(* IEC 61131-3 sources: 2026_Projet_YGO_ExcavatriceDragage/TOOLS/TEST_AUTO_CI/RESULTS/M_MAIN/reports, 9 files *)

(* ---- FB_CfgT330Normalizer_test.st ---- *)
(* =======================================================================
   🧪 FB_CfgT330Normalizer — cas ST unitaires du plan T330 (C3 v1.3)
   ───────────────────────────────────────────────────────────────
   Périmètre STRICT : le FB de normalisation des réglages HAUT, en boîte
   noire (contrat light : Enable / InHoming -> Ready / Corrected).
   Aucune assertion ne porte sur un consommateur (PRG_03 / PRG_04 /
   PRG_06 / GVL_PERSISTENT) : ces cas relèvent d'un lot d'intégration
   dédié (voir TASK_CONTRACT_T341, section « hors scope »).

   ── Conventions ───────────────────────────────────────────────────────
   1) 1 appel fb(...) = 1 scan.
   2) ⚠️ STruCpp v0.6.2 passe les VAR_IN_OUT par COPIE et ne génère que le
      copy-IN. La restitution `cfg := fb.CommunCfg;` est donc OBLIGATOIRE
      après chaque appel : elle émule la sémantique par RÉFÉRENCE de
      CODESYS. Sans elle, toute assertion de correction serait VACUE
      (le FB écrirait dans sa copie privée, jamais dans la variable de test).
      Le post-traitement `inject_var_in_out_copyout.py` ne s'applique PAS à
      une VAR déclarée dans un bloc `VAR` local de TEST (sa regex exige le
      préfixe `s.` que ce build n'émet pas) — d'où l'émulation explicite.
   3) ⚠️ Aucune assertion n'est placée dans une boucle FOR/WHILE : ce build
      STruCpp SUPPRIME silencieusement les ASSERT_* du corps d'une boucle
      (vérifié dans le C++ généré). Les balayages sont donc déroulés.
   4) Tolérance 1e-6 : les REAL sont en simple précision, un littéral ST est
      lu en double — un écart de ~1,4e-7 est normal sur 7,4999.
   5) Amorcage : le FB amorce ses mémoires de front au PREMIER scan où
      `Enable` est vrai, depuis les valeurs RESTAURÉES (piège P2 du cadrage).
      Une stimulation « saisie opérateur » se joue donc au scan SUIVANT.

   Référence : DOC/WFLOW/AUDITS/DESIGN/PLAN_T330_C3_INVARIANT_HAUT_v1.0.md §4.2
   ======================================================================= *)

SETUP
VAR
    FB       : FB_CfgT330Normalizer;
    WinchCfg : ST_WinchCfg;
    ComCfg   : ST_CommunCfg;
END_VAR
END_SETUP

(* ── Groupe A · Normalisation (TC-P10-056 .. TC-P10-062) ──────────────── *)

TEST 'TC-P10-056 R1 — FDC saisi trop haut : FDC corrige, TOP preserve'
VAR
    winchCfg  : ST_WinchCfg;
    communCfg : ST_CommunCfg;
END_VAR
    (* Scan 1 : amorcage sur la config restauree valide (8,50 / 7,50 / 0,50). *)
    winchCfg.CfgTopSensorPos_M := 8.5;
    communCfg.CfgCableLimitAscent_M := 7.5;
    communCfg.WinchSlowdownDistanceTop_M := 0.5;
    FB.Enable := TRUE;
    FB.InHoming := FALSE;
    FB(WinchCfgM1 := winchCfg, CommunCfg := communCfg);
    winchCfg := FB.WinchCfgM1;  communCfg := FB.CommunCfg;
    ASSERT_FALSE(FB.Corrected, 'Scan d amorcage : config valide, aucune correction');

    (* Scan 2 : l'operateur saisit FDC = 8,70 m (TOP inchange a 8,50 m). *)
    communCfg.CfgCableLimitAscent_M := 8.7;
    FB(WinchCfgM1 := winchCfg, CommunCfg := communCfg);
    winchCfg := FB.WinchCfgM1;  communCfg := FB.CommunCfg;
    ASSERT_NEAR(communCfg.CfgCableLimitAscent_M, 7.5, 0.000001,
                'R1 : FDC ramene a TOP - 1,00 m = 7,50');
    ASSERT_NEAR(winchCfg.CfgTopSensorPos_M, 8.5, 0.000001, 'R1 : le TOP n est PAS modifie');
    ASSERT_TRUE(FB.Corrected, 'R1 : une correction a eu lieu, message emis');
END_TEST

TEST 'TC-P10-057 R2 — TOP saisi trop bas : TOP corrige, FDC preserve'
VAR
    winchCfg  : ST_WinchCfg;
    communCfg : ST_CommunCfg;
END_VAR
    winchCfg.CfgTopSensorPos_M := 8.5;
    communCfg.CfgCableLimitAscent_M := 7.5;
    communCfg.WinchSlowdownDistanceTop_M := 0.5;
    FB.Enable := TRUE;
    FB.InHoming := FALSE;
    FB(WinchCfgM1 := winchCfg, CommunCfg := communCfg);
    winchCfg := FB.WinchCfgM1;  communCfg := FB.CommunCfg;

    (* Scan 2 : l'operateur saisit TOP = 7,00 m (FDC inchange a 7,50 m). *)
    winchCfg.CfgTopSensorPos_M := 7.0;
    FB(WinchCfgM1 := winchCfg, CommunCfg := communCfg);
    winchCfg := FB.WinchCfgM1;  communCfg := FB.CommunCfg;
    ASSERT_NEAR(winchCfg.CfgTopSensorPos_M, 8.5, 0.000001,
                'R2 : TOP ramene a FDC + 1,00 m = 8,50 (le champ saisi est corrige)');
    ASSERT_NEAR(communCfg.CfgCableLimitAscent_M, 7.5, 0.000001, 'R2 : le FDC n est PAS modifie');
    ASSERT_TRUE(FB.Corrected, 'R2 : une correction a eu lieu, message emis');
END_TEST

TEST 'TC-P10-058 R1 — Delta = 0,90 m : correction du champ saisi (FDC)'
VAR
    winchCfg  : ST_WinchCfg;
    communCfg : ST_CommunCfg;
END_VAR
    winchCfg.CfgTopSensorPos_M := 8.5;
    communCfg.CfgCableLimitAscent_M := 7.5;
    communCfg.WinchSlowdownDistanceTop_M := 0.5;
    FB.Enable := TRUE;
    FB.InHoming := FALSE;
    FB(WinchCfgM1 := winchCfg, CommunCfg := communCfg);
    winchCfg := FB.WinchCfgM1;  communCfg := FB.CommunCfg;

    (* Scan 2 : FDC = 7,60 m => Delta = 8,50 - 7,60 = 0,90 m < 1,00 m. *)
    communCfg.CfgCableLimitAscent_M := 7.6;
    FB(WinchCfgM1 := winchCfg, CommunCfg := communCfg);
    winchCfg := FB.WinchCfgM1;  communCfg := FB.CommunCfg;
    ASSERT_NEAR(communCfg.CfgCableLimitAscent_M, 7.5, 0.000001, 'Delta < 1,00 m : FDC ramene a 7,50');
    ASSERT_NEAR(winchCfg.CfgTopSensorPos_M, 8.5, 0.000001, 'Delta < 1,00 m : TOP preserve');
    ASSERT_TRUE(FB.Corrected, 'Delta < 1,00 m : correction signalee');
END_TEST

TEST 'TC-P10-059 R3 — plancher du ralentissement haut (0,20 -> 0,50)'
VAR
    winchCfg  : ST_WinchCfg;
    communCfg : ST_CommunCfg;
END_VAR
    winchCfg.CfgTopSensorPos_M := 8.5;
    communCfg.CfgCableLimitAscent_M := 7.5;
    communCfg.WinchSlowdownDistanceTop_M := 0.5;
    FB.Enable := TRUE;
    FB.InHoming := FALSE;
    FB(WinchCfgM1 := winchCfg, CommunCfg := communCfg);
    winchCfg := FB.WinchCfgM1;  communCfg := FB.CommunCfg;

    (* Scan 2 : ralentissement saisi a 0,20 m (< 0,50 m). *)
    communCfg.WinchSlowdownDistanceTop_M := 0.2;
    FB(WinchCfgM1 := winchCfg, CommunCfg := communCfg);
    winchCfg := FB.WinchCfgM1;  communCfg := FB.CommunCfg;
    ASSERT_NEAR(communCfg.WinchSlowdownDistanceTop_M, 0.5, 0.000001,
                'R3 : ralentissement ramene au plancher 0,50 m');
    ASSERT_NEAR(winchCfg.CfgTopSensorPos_M, 8.5, 0.000001, 'R3 : TOP inchange');
    ASSERT_NEAR(communCfg.CfgCableLimitAscent_M, 7.5, 0.000001, 'R3 : FDC inchange');
    ASSERT_TRUE(FB.Corrected, 'R3 : correction signalee');
END_TEST

TEST 'TC-P10-060 config valide (Delta = 2,50) : aucune correction, aucun message'
VAR
    winchCfg  : ST_WinchCfg;
    communCfg : ST_CommunCfg;
END_VAR
    winchCfg.CfgTopSensorPos_M := 8.5;
    communCfg.CfgCableLimitAscent_M := 7.5;
    communCfg.WinchSlowdownDistanceTop_M := 0.5;
    FB.Enable := TRUE;
    FB.InHoming := FALSE;
    FB(WinchCfgM1 := winchCfg, CommunCfg := communCfg);
    winchCfg := FB.WinchCfgM1;  communCfg := FB.CommunCfg;

    (* Scan 2 : TOP = 10,00 m, FDC = 7,50 m => Delta = 2,50 m, valide. *)
    winchCfg.CfgTopSensorPos_M := 10.0;
    FB(WinchCfgM1 := winchCfg, CommunCfg := communCfg);
    winchCfg := FB.WinchCfgM1;  communCfg := FB.CommunCfg;
    ASSERT_NEAR(winchCfg.CfgTopSensorPos_M, 10.0, 0.000001, 'Config valide : TOP preserve');
    ASSERT_NEAR(communCfg.CfgCableLimitAscent_M, 7.5, 0.000001, 'Config valide : FDC preserve');
    ASSERT_FALSE(FB.Corrected, 'Config valide : AUCUN message (compteur de messages = 0)');
END_TEST

TEST 'TC-P10-061 Q17 — les DEUX champs changent au meme scan : TOP preserve, FDC corrige'
VAR
    winchCfg  : ST_WinchCfg;
    communCfg : ST_CommunCfg;
END_VAR
    winchCfg.CfgTopSensorPos_M := 8.5;
    communCfg.CfgCableLimitAscent_M := 7.5;
    communCfg.WinchSlowdownDistanceTop_M := 0.5;
    FB.Enable := TRUE;
    FB.InHoming := FALSE;
    FB(WinchCfgM1 := winchCfg, CommunCfg := communCfg);
    winchCfg := FB.WinchCfgM1;  communCfg := FB.CommunCfg;

    (* Scan 2 : les 3 reglages changent ensemble : FDC 9,50 / TOP 8,00 / slowdown 0,10. *)
    communCfg.CfgCableLimitAscent_M := 9.5;
    winchCfg.CfgTopSensorPos_M := 8.0;
    communCfg.WinchSlowdownDistanceTop_M := 0.1;
    FB(WinchCfgM1 := winchCfg, CommunCfg := communCfg);
    winchCfg := FB.WinchCfgM1;  communCfg := FB.CommunCfg;
    ASSERT_NEAR(winchCfg.CfgTopSensorPos_M, 8.0, 0.000001, 'Q17 : le TOP saisi est PRESERVE');
    ASSERT_NEAR(communCfg.CfgCableLimitAscent_M, 7.0, 0.000001,
                'Q17 : FDC = TOP - 1,00 m = 7,00 (R0 a d abord ramene 9,50 a 9,00)');
    ASSERT_NEAR(communCfg.WinchSlowdownDistanceTop_M, 0.5, 0.000001, 'R3 : ralentissement ramene a 0,50');
    ASSERT_TRUE(FB.Corrected, 'Q17 : les trois corrections sont signalees');
END_TEST

TEST 'TC-P10-062 FDC = 0,00 m (borne basse, Delta valide) : accepte, aucune correction'
VAR
    winchCfg  : ST_WinchCfg;
    communCfg : ST_CommunCfg;
END_VAR
    winchCfg.CfgTopSensorPos_M := 8.5;
    communCfg.CfgCableLimitAscent_M := 7.5;
    communCfg.WinchSlowdownDistanceTop_M := 0.5;
    FB.Enable := TRUE;
    FB.InHoming := FALSE;
    FB(WinchCfgM1 := winchCfg, CommunCfg := communCfg);
    winchCfg := FB.WinchCfgM1;  communCfg := FB.CommunCfg;

    (* Scan 2 : FDC = 0,00 m => Delta = 8,50 m, valide. La borne basse est INCLUSE. *)
    communCfg.CfgCableLimitAscent_M := 0.0;
    FB(WinchCfgM1 := winchCfg, CommunCfg := communCfg);
    winchCfg := FB.WinchCfgM1;  communCfg := FB.CommunCfg;
    ASSERT_NEAR(communCfg.CfgCableLimitAscent_M, 0.0, 0.000001,
                'FDC a la borne basse : valeur ACCEPTEE telle quelle');
    ASSERT_NEAR(winchCfg.CfgTopSensorPos_M, 8.5, 0.000001, 'FDC a la borne basse : TOP inchange');
    ASSERT_FALSE(FB.Corrected, 'FDC a la borne basse : aucune correction, aucun message');
END_TEST

(* ── Groupe B · Idempotence et non-rebond (TC-P10-063 .. TC-P10-068) ──── *)

TEST 'TC-P10-063 Q24 — idempotence : le 2e scan apres correction ne corrige PLUS'
VAR
    winchCfg  : ST_WinchCfg;
    communCfg : ST_CommunCfg;
END_VAR
    winchCfg.CfgTopSensorPos_M := 8.5;
    communCfg.CfgCableLimitAscent_M := 7.5;
    communCfg.WinchSlowdownDistanceTop_M := 0.5;
    FB.Enable := TRUE;
    FB.InHoming := FALSE;
    FB(WinchCfgM1 := winchCfg, CommunCfg := communCfg);
    winchCfg := FB.WinchCfgM1;  communCfg := FB.CommunCfg;

    (* Scan 2 : correction (FDC 8,70 -> 7,50). *)
    communCfg.CfgCableLimitAscent_M := 8.7;
    FB(WinchCfgM1 := winchCfg, CommunCfg := communCfg);
    winchCfg := FB.WinchCfgM1;  communCfg := FB.CommunCfg;
    ASSERT_NEAR(communCfg.CfgCableLimitAscent_M, 7.5, 0.000001, 'Scan 2 : FDC corrige a 7,50');

    (* Scan 3 : rejeu SANS nouvelle saisie => ni correction, ni message, valeur stable. *)
    FB(WinchCfgM1 := winchCfg, CommunCfg := communCfg);
    winchCfg := FB.WinchCfgM1;  communCfg := FB.CommunCfg;
    ASSERT_NEAR(communCfg.CfgCableLimitAscent_M, 7.5, 0.000001, 'Scan 3 : valeur STABLE a 7,50');
    ASSERT_FALSE(FB.Corrected, 'Scan 3 : AUCUNE seconde correction (test probatoire de Q24)');
END_TEST

TEST 'TC-P10-064 reserve EXACTEMENT 1,00 m : aucune correction (aucun epsilon)'
VAR
    winchCfg  : ST_WinchCfg;
    communCfg : ST_CommunCfg;
END_VAR
    winchCfg.CfgTopSensorPos_M := 8.5;
    communCfg.CfgCableLimitAscent_M := 7.5;
    communCfg.WinchSlowdownDistanceTop_M := 0.5;
    FB.Enable := TRUE;
    FB.InHoming := FALSE;
    FB(WinchCfgM1 := winchCfg, CommunCfg := communCfg);
    winchCfg := FB.WinchCfgM1;  communCfg := FB.CommunCfg;
    ASSERT_FALSE(FB.Corrected, 'Delta = 1,00 m exactement : aucune correction (comparaison stricte)');
    ASSERT_NEAR(winchCfg.CfgTopSensorPos_M - communCfg.CfgCableLimitAscent_M, 1.0, 0.000001,
                'Le flottant est EXACT : 8,50 - 7,50 = 1,00 (aucun eps necessaire)');

    (* Scan 2 : rejeu identique — la reserve reste exactement 1,00 m. *)
    FB(WinchCfgM1 := winchCfg, CommunCfg := communCfg);
    winchCfg := FB.WinchCfgM1;  communCfg := FB.CommunCfg;
    ASSERT_FALSE(FB.Corrected, 'Scan 2 : aucune oscillation autour du seuil');
END_TEST

TEST 'TC-P10-065 pt1 balayage 7,4999 — Delta = 1,0001 m : FDC conserve'
VAR
    winchCfg  : ST_WinchCfg;
    communCfg : ST_CommunCfg;
END_VAR
    winchCfg.CfgTopSensorPos_M := 8.5;
    communCfg.CfgCableLimitAscent_M := 7.5;
    communCfg.WinchSlowdownDistanceTop_M := 0.5;
    FB.Enable := TRUE;
    FB.InHoming := FALSE;
    FB(WinchCfgM1 := winchCfg, CommunCfg := communCfg);
    winchCfg := FB.WinchCfgM1;  communCfg := FB.CommunCfg;

    communCfg.CfgCableLimitAscent_M := 7.4999;
    FB(WinchCfgM1 := winchCfg, CommunCfg := communCfg);
    winchCfg := FB.WinchCfgM1;  communCfg := FB.CommunCfg;
    ASSERT_NEAR(communCfg.CfgCableLimitAscent_M, 7.4999, 0.000001,
                'Delta > 1,00 m : FDC conserve tel quel');
    ASSERT_FALSE(FB.Corrected, 'Delta > 1,00 m : aucun message');
END_TEST

TEST 'TC-P10-065 pt2 balayage 7,5000 — Delta = 1,00 m exactement : FDC conserve'
VAR
    winchCfg  : ST_WinchCfg;
    communCfg : ST_CommunCfg;
END_VAR
    winchCfg.CfgTopSensorPos_M := 8.5;
    communCfg.CfgCableLimitAscent_M := 7.5;
    communCfg.WinchSlowdownDistanceTop_M := 0.5;
    FB.Enable := TRUE;
    FB.InHoming := FALSE;
    FB(WinchCfgM1 := winchCfg, CommunCfg := communCfg);
    winchCfg := FB.WinchCfgM1;  communCfg := FB.CommunCfg;

    communCfg.CfgCableLimitAscent_M := 7.5;
    FB(WinchCfgM1 := winchCfg, CommunCfg := communCfg);
    winchCfg := FB.WinchCfgM1;  communCfg := FB.CommunCfg;
    ASSERT_NEAR(communCfg.CfgCableLimitAscent_M, 7.5, 0.000001,
                'Delta = 1,00 m (point limite INCLUS) : FDC conserve');
    ASSERT_FALSE(FB.Corrected, 'Delta = 1,00 m : aucun message');
END_TEST

TEST 'TC-P10-065 pt3 balayage 7,5001 — Delta = 0,9999 m : FDC corrige, une seule fois'
VAR
    winchCfg  : ST_WinchCfg;
    communCfg : ST_CommunCfg;
END_VAR
    winchCfg.CfgTopSensorPos_M := 8.5;
    communCfg.CfgCableLimitAscent_M := 7.5;
    communCfg.WinchSlowdownDistanceTop_M := 0.5;
    FB.Enable := TRUE;
    FB.InHoming := FALSE;
    FB(WinchCfgM1 := winchCfg, CommunCfg := communCfg);
    winchCfg := FB.WinchCfgM1;  communCfg := FB.CommunCfg;

    communCfg.CfgCableLimitAscent_M := 7.5001;
    FB(WinchCfgM1 := winchCfg, CommunCfg := communCfg);
    winchCfg := FB.WinchCfgM1;  communCfg := FB.CommunCfg;
    ASSERT_NEAR(communCfg.CfgCableLimitAscent_M, 7.5, 0.000001, 'Delta < 1,00 m : FDC ramene a 7,50');
    ASSERT_TRUE(FB.Corrected, 'Delta < 1,00 m : correction signalee');

    (* Scan suivant : la valeur corrigee ne rebondit pas (aucune oscillation au seuil). *)
    FB(WinchCfgM1 := winchCfg, CommunCfg := communCfg);
    winchCfg := FB.WinchCfgM1;  communCfg := FB.CommunCfg;
    ASSERT_FALSE(FB.Corrected, 'Scan suivant : aucune seconde correction (pas d oscillation)');
END_TEST

TEST 'TC-P10-066 LIMITE DECLAREE — guerre d ecriture IHM : correction a CHAQUE scan'
VAR
    winchCfg  : ST_WinchCfg;
    communCfg : ST_CommunCfg;
END_VAR
    (* ⚠️ Ce cas fige une LIMITE ASSUMEE du lot (plan v1.3 §4.2, C3), PAS une exigence :
       si le panneau IHM reecrit 8,70 m a CHAQUE scan, la normalisation corrige a chaque
       scan et le message rebondit — aucun amortissement n'est specifie ni implemente.
       Le test est volontairement falsifiable : ajouter un anti-rebond le fera echouer,
       ce qui forcera une decision DOCUMENTEE plutot qu'une derive silencieuse.
       Balayage DEROULE (3 scans) : une assertion dans une boucle serait supprimee
       silencieusement par STruCpp et le test deviendrait VACUE. *)
    winchCfg.CfgTopSensorPos_M := 8.5;
    communCfg.CfgCableLimitAscent_M := 7.5;
    communCfg.WinchSlowdownDistanceTop_M := 0.5;
    FB.Enable := TRUE;
    FB.InHoming := FALSE;
    FB(WinchCfgM1 := winchCfg, CommunCfg := communCfg);
    winchCfg := FB.WinchCfgM1;  communCfg := FB.CommunCfg;

    (* Scan 2. *)
    communCfg.CfgCableLimitAscent_M := 8.7;
    FB(WinchCfgM1 := winchCfg, CommunCfg := communCfg);
    winchCfg := FB.WinchCfgM1;  communCfg := FB.CommunCfg;
    ASSERT_NEAR(communCfg.CfgCableLimitAscent_M, 7.5, 0.000001, 'Scan 2 : correction reappliquee');
    ASSERT_TRUE(FB.Corrected, 'Scan 2 : message emis (rebond ASSUME)');

    (* Scan 3. *)
    communCfg.CfgCableLimitAscent_M := 8.7;
    FB(WinchCfgM1 := winchCfg, CommunCfg := communCfg);
    winchCfg := FB.WinchCfgM1;  communCfg := FB.CommunCfg;
    ASSERT_NEAR(communCfg.CfgCableLimitAscent_M, 7.5, 0.000001, 'Scan 3 : correction reappliquee');
    ASSERT_TRUE(FB.Corrected, 'Scan 3 : message emis (rebond ASSUME)');

    (* Scan 4. *)
    communCfg.CfgCableLimitAscent_M := 8.7;
    FB(WinchCfgM1 := winchCfg, CommunCfg := communCfg);
    winchCfg := FB.WinchCfgM1;  communCfg := FB.CommunCfg;
    ASSERT_NEAR(communCfg.CfgCableLimitAscent_M, 7.5, 0.000001, 'Scan 4 : correction reappliquee');
    ASSERT_TRUE(FB.Corrected, 'Scan 4 : message emis (rebond ASSUME)');
END_TEST

TEST 'TC-P10-067 valeur IDENTIQUE re-saisie : aucun front, aucune correction'
VAR
    winchCfg  : ST_WinchCfg;
    communCfg : ST_CommunCfg;
END_VAR
    winchCfg.CfgTopSensorPos_M := 8.5;
    communCfg.CfgCableLimitAscent_M := 7.5;
    communCfg.WinchSlowdownDistanceTop_M := 0.5;
    FB.Enable := TRUE;
    FB.InHoming := FALSE;
    FB(WinchCfgM1 := winchCfg, CommunCfg := communCfg);
    winchCfg := FB.WinchCfgM1;  communCfg := FB.CommunCfg;

    (* Scan 2 : le champ est REEcrit avec la MEME valeur (8,50 -> 8,50). *)
    winchCfg.CfgTopSensorPos_M := 8.5;
    FB(WinchCfgM1 := winchCfg, CommunCfg := communCfg);
    winchCfg := FB.WinchCfgM1;  communCfg := FB.CommunCfg;
    ASSERT_FALSE(FB.Corrected, 'Valeur identique re-saisie : aucun front, aucun message');
    ASSERT_NEAR(winchCfg.CfgTopSensorPos_M, 8.5, 0.000001, 'Valeur identique : TOP inchange');
END_TEST

TEST 'TC-P10-068 changement de page IHM sans modification : aucune correction'
VAR
    winchCfg  : ST_WinchCfg;
    communCfg : ST_CommunCfg;
END_VAR
    winchCfg.CfgTopSensorPos_M := 8.5;
    communCfg.CfgCableLimitAscent_M := 7.5;
    communCfg.WinchSlowdownDistanceTop_M := 0.5;
    FB.Enable := TRUE;
    FB.InHoming := FALSE;
    FB(WinchCfgM1 := winchCfg, CommunCfg := communCfg);
    winchCfg := FB.WinchCfgM1;  communCfg := FB.CommunCfg;

    (* Scan 2 : page quittee => normalisation suspendue, AUCUNE valeur modifiee. *)
    FB.Enable := FALSE;
    FB(WinchCfgM1 := winchCfg, CommunCfg := communCfg);
    winchCfg := FB.WinchCfgM1;  communCfg := FB.CommunCfg;
    ASSERT_FALSE(FB.Corrected, 'Normalisation suspendue : aucun message');
    ASSERT_FALSE(FB.Ready, 'Normalisation suspendue : Ready = FALSE');

    (* Scan 3 : retour sur la page, valeurs inchangees => ni front, ni correction. *)
    FB.Enable := TRUE;
    FB(WinchCfgM1 := winchCfg, CommunCfg := communCfg);
    winchCfg := FB.WinchCfgM1;  communCfg := FB.CommunCfg;
    ASSERT_FALSE(FB.Corrected, 'Retour de page sans modification : aucune correction');
    ASSERT_NEAR(winchCfg.CfgTopSensorPos_M, 8.5, 0.000001, 'Retour de page : TOP inchange');
    ASSERT_NEAR(communCfg.CfgCableLimitAscent_M, 7.5, 0.000001, 'Retour de page : FDC inchange');
END_TEST

(* ── Groupe C · Boot, restauration, hot restart (TC-P10-069 .. TC-P10-074) ─ *)

TEST 'TC-P10-069 NVRAM valide au demarrage a froid : 0 correction, valeurs preservees'
VAR
    winchCfg  : ST_WinchCfg;
    communCfg : ST_CommunCfg;
END_VAR
    winchCfg.CfgTopSensorPos_M := 8.5;
    communCfg.CfgCableLimitAscent_M := 7.5;
    communCfg.WinchSlowdownDistanceTop_M := 0.5;
    FB.Enable := TRUE;
    FB.InHoming := FALSE;
    FB(WinchCfgM1 := winchCfg, CommunCfg := communCfg);
    winchCfg := FB.WinchCfgM1;  communCfg := FB.CommunCfg;
    ASSERT_TRUE(FB.Ready, 'Normalisation ARMED des le premier scan apres restauration');
    ASSERT_FALSE(FB.Corrected, 'NVRAM valide : aucune correction');
    ASSERT_NEAR(winchCfg.CfgTopSensorPos_M, 8.5, 0.000001, 'NVRAM valide : TOP preserve');
    ASSERT_NEAR(communCfg.CfgCableLimitAscent_M, 7.5, 0.000001, 'NVRAM valide : FDC preserve');
    ASSERT_NEAR(communCfg.WinchSlowdownDistanceTop_M, 0.5, 0.000001, 'NVRAM valide : ralentissement preserve');
END_TEST

TEST 'TC-P10-070 NVRAM invalide au demarrage a froid : Q17 (TOP preserve, FDC corrige)'
VAR
    winchCfg  : ST_WinchCfg;
    communCfg : ST_CommunCfg;
END_VAR
    (* NVRAM restauree INVALIDE : TOP = 7,00 m / FDC = 7,50 m. *)
    winchCfg.CfgTopSensorPos_M := 7.0;
    communCfg.CfgCableLimitAscent_M := 7.5;
    communCfg.WinchSlowdownDistanceTop_M := 0.5;
    FB.Enable := TRUE;
    FB.InHoming := FALSE;
    FB(WinchCfgM1 := winchCfg, CommunCfg := communCfg);
    winchCfg := FB.WinchCfgM1;  communCfg := FB.CommunCfg;
    ASSERT_NEAR(winchCfg.CfgTopSensorPos_M, 7.0, 0.000001,
                'Q17 : le TOP restaure est PRESERVE (c est la cote gravee par le homing)');
    ASSERT_NEAR(communCfg.CfgCableLimitAscent_M, 6.0, 0.000001, 'Q17 : FDC = TOP - 1,00 m = 6,00');
    ASSERT_TRUE(FB.Corrected, 'NVRAM invalide : correction signalee');
END_TEST

TEST 'TC-P10-071 premier scan NOT Initialized : normalisation INHIBEE, aucune ecriture'
VAR
    winchCfg  : ST_WinchCfg;
    communCfg : ST_CommunCfg;
END_VAR
    (* Ponts non restaures : les valeurs presentes sont les DEFAUTS DUT, pas une saisie. *)
    winchCfg.CfgTopSensorPos_M := 99.0;
    communCfg.CfgCableLimitAscent_M := 99.0;
    communCfg.WinchSlowdownDistanceTop_M := 99.0;
    FB.Enable := FALSE;
    FB.InHoming := FALSE;
    FB(WinchCfgM1 := winchCfg, CommunCfg := communCfg);
    winchCfg := FB.WinchCfgM1;  communCfg := FB.CommunCfg;
    ASSERT_FALSE(FB.Ready, 'NOT Initialized : normalisation NON armee');
    ASSERT_FALSE(FB.Corrected, 'NOT Initialized : aucun message');
    ASSERT_NEAR(winchCfg.CfgTopSensorPos_M, 99.0, 0.000001, 'NOT Initialized : AUCUNE ecriture TOP');
    ASSERT_NEAR(communCfg.CfgCableLimitAscent_M, 99.0, 0.000001, 'NOT Initialized : AUCUNE ecriture FDC');
    ASSERT_NEAR(communCfg.WinchSlowdownDistanceTop_M, 99.0, 0.000001,
                'NOT Initialized : AUCUNE ecriture ralentissement');
END_TEST

TEST 'TC-P10-074 ptA restauration NVRAM : AUCUNE correction fantome (defauts DUT -> restaure)'
VAR
    winchCfg  : ST_WinchCfg;
    communCfg : ST_CommunCfg;
END_VAR
    (* PREUVE EXIGEE par le plan §2.2 point 3 : la transition « defauts DUT ->
       valeurs RESTAUREES » ne doit PAS etre prise pour une saisie operateur. *)
    winchCfg.CfgTopSensorPos_M := 8.5;      (* defauts DUT au 1er scan *)
    communCfg.CfgCableLimitAscent_M := 7.5;
    communCfg.WinchSlowdownDistanceTop_M := 0.5;
    FB.Enable := FALSE;                     (* ponts non restaures *)
    FB.InHoming := FALSE;
    FB(WinchCfgM1 := winchCfg, CommunCfg := communCfg);
    winchCfg := FB.WinchCfgM1;  communCfg := FB.CommunCfg;

    winchCfg.CfgTopSensorPos_M := 8.5;      (* valeurs RESTAUREES, valides *)
    communCfg.CfgCableLimitAscent_M := 7.5;
    communCfg.WinchSlowdownDistanceTop_M := 0.5;
    FB.Enable := TRUE;
    FB(WinchCfgM1 := winchCfg, CommunCfg := communCfg);
    winchCfg := FB.WinchCfgM1;  communCfg := FB.CommunCfg;
    ASSERT_FALSE(FB.Corrected, 'Restauration NVRAM : AUCUNE correction fantome');
    ASSERT_NEAR(winchCfg.CfgTopSensorPos_M, 8.5, 0.000001, 'Restauration NVRAM : TOP preserve');
    ASSERT_NEAR(communCfg.CfgCableLimitAscent_M, 7.5, 0.000001, 'Restauration NVRAM : FDC preserve');
END_TEST

TEST 'TC-P10-074 ptB download/RTS : comportement DETERMINISTE, une seule correction'
VAR
    winchCfg  : ST_WinchCfg;
    communCfg : ST_CommunCfg;
END_VAR
    (* NVRAM restauree INVALIDE apres download : une correction, jamais repetee. *)
    winchCfg.CfgTopSensorPos_M := 7.0;
    communCfg.CfgCableLimitAscent_M := 7.5;
    communCfg.WinchSlowdownDistanceTop_M := 0.5;
    FB.Enable := TRUE;
    FB.InHoming := FALSE;
    FB(WinchCfgM1 := winchCfg, CommunCfg := communCfg);
    winchCfg := FB.WinchCfgM1;  communCfg := FB.CommunCfg;
    ASSERT_TRUE(FB.Corrected, 'NVRAM invalide : une correction, signalee');
    ASSERT_NEAR(communCfg.CfgCableLimitAscent_M, 6.0, 0.000001, 'NVRAM invalide : FDC = 6,00 (Q17)');

    FB(WinchCfgM1 := winchCfg, CommunCfg := communCfg);
    winchCfg := FB.WinchCfgM1;  communCfg := FB.CommunCfg;
    ASSERT_FALSE(FB.Corrected, 'Scan suivant : aucune correction fantome repetee');
    ASSERT_NEAR(communCfg.CfgCableLimitAscent_M, 6.0, 0.000001, 'Valeur corrigee STABLE');
END_TEST

(* ── Groupe E · Modes et domaines (TC-P10-082 .. TC-P10-092) ──────────── *)

TEST 'TC-P10-082 Q22/C2 — homing : gel NVRAM, repli NIVEAU Q17, non-memorisation'
VAR
    winchCfg  : ST_WinchCfg;
    communCfg : ST_CommunCfg;
    fbRestart : FB_CfgT330Normalizer;
    wR        : ST_WinchCfg;
    cR        : ST_CommunCfg;
END_VAR
    (* Scan 1 : config valide, hors homing. *)
    winchCfg.CfgTopSensorPos_M := 8.5;
    communCfg.CfgCableLimitAscent_M := 7.5;
    communCfg.WinchSlowdownDistanceTop_M := 0.5;
    FB.Enable := TRUE;
    FB.InHoming := FALSE;
    FB(WinchCfgM1 := winchCfg, CommunCfg := communCfg);
    winchCfg := FB.WinchCfgM1;  communCfg := FB.CommunCfg;

    (* ① PENDANT le homing : TOP saisi 7,00 m => R2 INHIBEE et NVRAM GELEE (aucune ecriture). *)
    winchCfg.CfgTopSensorPos_M := 7.0;
    FB.InHoming := TRUE;
    FB(WinchCfgM1 := winchCfg, CommunCfg := communCfg);
    winchCfg := FB.WinchCfgM1;  communCfg := FB.CommunCfg;
    ASSERT_NEAR(winchCfg.CfgTopSensorPos_M, 7.0, 0.000001,
                'Homing : le TOP saisi reste 7,00 INCHANGE (R2 inhibee, gel NVRAM)');
    ASSERT_NEAR(communCfg.CfgCableLimitAscent_M, 7.5, 0.000001, 'Homing : FDC gele');
    ASSERT_FALSE(FB.Corrected, 'Homing : aucune ecriture Cfg, donc aucun message');

    (* ② SORTIE du homing : la config est toujours invalide => REPLI NIVEAU = Q17. *)
    FB.InHoming := FALSE;
    FB(WinchCfgM1 := winchCfg, CommunCfg := communCfg);
    winchCfg := FB.WinchCfgM1;  communCfg := FB.CommunCfg;
    ASSERT_NEAR(winchCfg.CfgTopSensorPos_M, 7.0, 0.000001, 'Sortie de homing : TOP PRESERVE (Q17)');
    ASSERT_NEAR(communCfg.CfgCableLimitAscent_M, 6.0, 0.000001,
                'Sortie de homing : FDC = 7,00 - 1,00 = 6,00 (repli NIVEAU)');
    ASSERT_TRUE(FB.Corrected, 'Sortie de homing : message NOMINAL, une seule fois');

    (* ③ Scan suivant : AUCUNE seconde correction (idempotence). *)
    FB(WinchCfgM1 := winchCfg, CommunCfg := communCfg);
    winchCfg := FB.WinchCfgM1;  communCfg := FB.CommunCfg;
    ASSERT_FALSE(FB.Corrected, 'Scan suivant : aucune seconde correction');
    ASSERT_NEAR(communCfg.CfgCableLimitAscent_M, 6.0, 0.000001, 'Scan suivant : FDC stable a 6,00');

    (* ④ Variante (c) — coupure pendant le homing : l intention est PERDUE. Un redemarrage
       a froid (instance NEUVE : les memoires du FB ne sont pas persistantes) applique la
       normalisation Q2 ORDINAIRE : rien de specifique n a ete memorise. *)
    wR.CfgTopSensorPos_M := 7.0;
    cR.CfgCableLimitAscent_M := 7.5;
    cR.WinchSlowdownDistanceTop_M := 0.5;
    fbRestart.Enable := TRUE;
    fbRestart.InHoming := FALSE;
    fbRestart(WinchCfgM1 := wR, CommunCfg := cR);
    wR := fbRestart.WinchCfgM1;  cR := fbRestart.CommunCfg;
    ASSERT_NEAR(wR.CfgTopSensorPos_M, 7.0, 0.000001, 'Redemarrage : TOP restaure preserve');
    ASSERT_NEAR(cR.CfgCableLimitAscent_M, 6.0, 0.000001, 'Redemarrage : Q2 ordinaire => FDC = 6,00');
    ASSERT_TRUE(fbRestart.Corrected, 'Redemarrage : message Q2 ordinaire (aucune memoire d intention)');
END_TEST

TEST 'TC-P10-090 ptA R0 — FDC = 0,00 m : valeur A LA BORNE, acceptee sans message'
VAR
    winchCfg  : ST_WinchCfg;
    communCfg : ST_CommunCfg;
END_VAR
    winchCfg.CfgTopSensorPos_M := 8.5;
    communCfg.CfgCableLimitAscent_M := 0.0;
    communCfg.WinchSlowdownDistanceTop_M := 0.5;
    FB.Enable := TRUE;
    FB.InHoming := FALSE;
    FB(WinchCfgM1 := winchCfg, CommunCfg := communCfg);
    winchCfg := FB.WinchCfgM1;  communCfg := FB.CommunCfg;
    ASSERT_NEAR(communCfg.CfgCableLimitAscent_M, 0.0, 0.000001, 'R0 : 0,00 m reste 0,00 m (borne INCLUSE)');
    ASSERT_FALSE(FB.Corrected, 'R0 : a la borne, aucune correction, aucun message');
END_TEST

TEST 'TC-P10-090 ptB R0 — FDC = -1,00 m : CLAMPE a 0,00 m + message'
VAR
    winchCfg  : ST_WinchCfg;
    communCfg : ST_CommunCfg;
END_VAR
    winchCfg.CfgTopSensorPos_M := 8.5;
    communCfg.CfgCableLimitAscent_M := -1.0;
    communCfg.WinchSlowdownDistanceTop_M := 0.5;
    FB.Enable := TRUE;
    FB.InHoming := FALSE;
    FB(WinchCfgM1 := winchCfg, CommunCfg := communCfg);
    winchCfg := FB.WinchCfgM1;  communCfg := FB.CommunCfg;
    ASSERT_NEAR(communCfg.CfgCableLimitAscent_M, 0.0, 0.000001, 'R0 : -1,00 m CLAMPE a 0,00 m');
    ASSERT_NEAR(winchCfg.CfgTopSensorPos_M, 8.5, 0.000001, 'R0 : TOP inchange (Delta = 8,50 m valide)');
    ASSERT_TRUE(FB.Corrected, 'R0 : clamp signale (jamais muet)');
END_TEST

TEST 'TC-P10-090 ptC R0 — TOP = 0,50 m : CLAMPE a 1,00 m + message, R0 observe SEUL'
VAR
    winchCfg  : ST_WinchCfg;
    communCfg : ST_CommunCfg;
END_VAR
    (* FDC = 0,00 m : apres clamp du TOP a 1,00 m, Delta = 1,00 m exactement => la regle
       Delta reste INERTE, ce qui isole R0 (exigence Q21 bis). *)
    winchCfg.CfgTopSensorPos_M := 0.5;
    communCfg.CfgCableLimitAscent_M := 0.0;
    communCfg.WinchSlowdownDistanceTop_M := 0.5;
    FB.Enable := TRUE;
    FB.InHoming := FALSE;
    FB(WinchCfgM1 := winchCfg, CommunCfg := communCfg);
    winchCfg := FB.WinchCfgM1;  communCfg := FB.CommunCfg;
    ASSERT_NEAR(winchCfg.CfgTopSensorPos_M, 1.0, 0.000001, 'R0 : TOP 0,50 m CLAMPE a 1,00 m');
    ASSERT_NEAR(communCfg.CfgCableLimitAscent_M, 0.0, 0.000001, 'R0 : FDC inchange a 0,00 m');
    ASSERT_TRUE(FB.Corrected, 'R0 : clamp signale (jamais muet)');
END_TEST

TEST 'TC-P10-091 ptA Q21 bis — R0 SEUL : Delta >= 1 avant clamp (FDC 9,50 / TOP 12,00)'
VAR
    winchCfg  : ST_WinchCfg;
    communCfg : ST_CommunCfg;
END_VAR
    (* LE cas probatoire : Delta = 2,50 m >= 1,00 m, donc AUCUNE regle Delta ne se
       declenche : SEUL R0 agit. Sans R0 en amont, ces deux valeurs restaient hors
       domaine indefiniment. *)
    winchCfg.CfgTopSensorPos_M := 12.0;
    communCfg.CfgCableLimitAscent_M := 9.5;
    communCfg.WinchSlowdownDistanceTop_M := 0.5;
    FB.Enable := TRUE;
    FB.InHoming := FALSE;
    FB(WinchCfgM1 := winchCfg, CommunCfg := communCfg);
    winchCfg := FB.WinchCfgM1;  communCfg := FB.CommunCfg;
    ASSERT_NEAR(communCfg.CfgCableLimitAscent_M, 9.0, 0.000001, 'Q21 bis : FDC ramene a la borne haute 9,00 m');
    ASSERT_NEAR(winchCfg.CfgTopSensorPos_M, 10.0, 0.000001, 'Q21 bis : TOP ramene a la borne haute 10,00 m');
    ASSERT_NEAR(winchCfg.CfgTopSensorPos_M - communCfg.CfgCableLimitAscent_M, 1.0, 0.000001,
                'Q21 bis : coherence Delta = 1,00 m APRES clamp');
    ASSERT_TRUE(FB.Corrected, 'Q21 bis : clamp signale, message non alarmant');
END_TEST

TEST 'TC-P10-091 ptB Q21 bis — domaines absurdes : R0 borne AVANT tout usage aval'
VAR
    winchCfg  : ST_WinchCfg;
    communCfg : ST_CommunCfg;
END_VAR
    winchCfg.CfgTopSensorPos_M := 150.0;
    communCfg.CfgCableLimitAscent_M := -150.0;
    communCfg.WinchSlowdownDistanceTop_M := 0.5;
    FB.Enable := TRUE;
    FB.InHoming := FALSE;
    FB(WinchCfgM1 := winchCfg, CommunCfg := communCfg);
    winchCfg := FB.WinchCfgM1;  communCfg := FB.CommunCfg;
    ASSERT_NEAR(communCfg.CfgCableLimitAscent_M, 0.0, 0.000001, 'Domaines absurdes : FDC borne a 0,00 m');
    ASSERT_NEAR(winchCfg.CfgTopSensorPos_M, 10.0, 0.000001, 'Domaines absurdes : TOP borne a 10,00 m');
    ASSERT_TRUE(winchCfg.CfgTopSensorPos_M <= 10.0, 'Aucune valeur hors domaine ne subsiste');
    ASSERT_TRUE(FB.Corrected, 'Domaines absurdes : clamp signale');
END_TEST

TEST 'TC-P10-092 ptA C1 — R0 d abord : TOP 11,00 -> 10,00 et FDC 10,00 -> 9,00, Delta valid'
VAR
    winchCfg  : ST_WinchCfg;
    communCfg : ST_CommunCfg;
END_VAR
    (* TOP volontairement AU-DELA de la borne : c'est ce qui rend le cas DISCRIMINANT.
       Si R0 ne s'appliquait pas, Delta = 11,00 - 10,00 = 1,00 m serait deja « valide »
       et AUCUNE regle ne corrigerait : les deux valeurs resteraient hors domaine.
       Avec R0 en amont : TOP -> 10,00, FDC -> 9,00, Delta final = 1,00 m exactement. *)
    winchCfg.CfgTopSensorPos_M := 11.0;
    communCfg.CfgCableLimitAscent_M := 10.0;
    communCfg.WinchSlowdownDistanceTop_M := 0.5;
    FB.Enable := TRUE;
    FB.InHoming := FALSE;
    FB(WinchCfgM1 := winchCfg, CommunCfg := communCfg);
    winchCfg := FB.WinchCfgM1;  communCfg := FB.CommunCfg;
    ASSERT_NEAR(communCfg.CfgCableLimitAscent_M, 9.0, 0.000001, 'C1 : FDC 10,00 m ramene a la borne 9,00 m');
    ASSERT_NEAR(winchCfg.CfgTopSensorPos_M, 10.0, 0.000001, 'C1 : TOP 11,00 m ramene a la borne 10,00 m');
    ASSERT_NEAR(winchCfg.CfgTopSensorPos_M - communCfg.CfgCableLimitAscent_M, 1.0, 0.000001,
                'C1 : Delta = 1,00 m exactement => aucune correction supplementaire');
    ASSERT_TRUE(FB.Corrected, 'C1 : seule la correction R0 est signalee');
END_TEST

TEST 'TC-P10-092 ptB C1 — R2 au plus haut de sa plage : TOP = 10,00 m, jamais au-dela'
VAR
    winchCfg  : ST_WinchCfg;
    communCfg : ST_CommunCfg;
END_VAR
    (* Amorcage a la borne haute : FDC = 9,00 m (borne), TOP = 10,00 m (Delta = 1,00 m). *)
    winchCfg.CfgTopSensorPos_M := 10.0;
    communCfg.CfgCableLimitAscent_M := 9.0;
    communCfg.WinchSlowdownDistanceTop_M := 0.5;
    FB.Enable := TRUE;
    FB.InHoming := FALSE;
    FB(WinchCfgM1 := winchCfg, CommunCfg := communCfg);
    winchCfg := FB.WinchCfgM1;  communCfg := FB.CommunCfg;
    ASSERT_FALSE(FB.Corrected, 'Amorcage a la borne haute : aucune correction');

    (* L'operateur saisit TOP = 2,00 m : R2 doit redonner EXACTEMENT 10,00 m. *)
    winchCfg.CfgTopSensorPos_M := 2.0;
    FB(WinchCfgM1 := winchCfg, CommunCfg := communCfg);
    winchCfg := FB.WinchCfgM1;  communCfg := FB.CommunCfg;
    ASSERT_NEAR(winchCfg.CfgTopSensorPos_M, 10.0, 0.000001,
                'C1 : R2 redonne exactement TOP = 10,00 m (jamais > 10,00)');
    ASSERT_TRUE(winchCfg.CfgTopSensorPos_M <= 10.0, 'C1 : aucune valeur hors borne ne peut etre produite');
    ASSERT_TRUE(FB.Corrected, 'C1 : correction signalee');
END_TEST

(* ---- MAIN_GLOBAL_test.st ---- *)
SETUP
VAR
    mainMachine : FB_Main_EndToEnd;
    stepBefore  : E_AutoCycleStep;   // mémoire étape séquenceur pour test relâchement homme-mort
END_VAR
END_SETUP

TEST 'MAIN_GLOBAL : Chaine Complete - Qualification Neutre vers Montee Treuils Couples'
    // 1. Initialisation boot au neutre (Raw = 5000)
    mainMachine(
        JoyRawX := 5000,
        JoyRawY := 5000,
        JoyDeadmanBtn := FALSE,
        CmdMode := E_Mode.MAINT_N1,
        CmdWinchSelect := 1,
        EmergencyChainClosed := TRUE,
        PowerContactorEngaged := TRUE
    );
    mainMachine(
        JoyRawX := 5000,
        JoyRawY := 5000,
        JoyDeadmanBtn := TRUE, // Début appui homme-mort au neutre
        CmdMode := E_Mode.MAINT_N1,
        CmdWinchSelect := 1,
        EmergencyChainClosed := TRUE,
        PowerContactorEngaged := TRUE
    );
    ADVANCE_TIME(150000000); // 150 ms (> 100 ms DeadmanArmHoldTime)
    mainMachine(
        JoyRawX := 5000,
        JoyRawY := 5000,
        JoyDeadmanBtn := TRUE, // Confirmation maintien homme-mort -> Armé
        CmdMode := E_Mode.MAINT_N1,
        CmdWinchSelect := 1,
        EmergencyChainClosed := TRUE,
        PowerContactorEngaged := TRUE
    );

    // 2. Stimulus Opérateur : Poussée Manche vers le Haut (+Y = 8000) avec Homme-mort maintenu
    mainMachine(
        JoyRawX := 5000,
        JoyRawY := 8000, // Déviation Y Montée
        JoyDeadmanBtn := TRUE,
        CmdMode := E_Mode.MAINT_N1,
        CmdWinchSelect := 1,
        EmergencyChainClosed := TRUE,
        PowerContactorEngaged := TRUE
    );
    mainMachine(
        JoyRawX := 5000,
        JoyRawY := 8000,
        JoyDeadmanBtn := TRUE,
        CmdMode := E_Mode.MAINT_N1,
        CmdWinchSelect := 1,
        EmergencyChainClosed := TRUE,
        PowerContactorEngaged := TRUE
    );

    // 3. Vérification des flux à travers toute la machine (PRG_02 -> PRG_07)
    // - Bus PRG_02 : Joystick armé et qualifié
    ASSERT_TRUE(mainMachine.BusAcq.Joystick.DeadmanArmed, 'PRG_02: Homme-mort qualifie');

    // - Bus PRG_03 : Mode Manuel N1 arbitré
    ASSERT_EQ(mainMachine.BusModes.Mode, E_Mode.MAINT_N1, 'PRG_03: Mode MAINT_N1 arbitre');

    // - Bus PRG_04 : Demande de montée et sécurité nominale
    ASSERT_FALSE(mainMachine.BusWinch.WinchM1Safety.SafeStop, 'PRG_04: Aucun SafeStop actif');

    // - Bus PRG_07 : Bandeau IHM informé sans défaut
    ASSERT_TRUE(mainMachine.BusBanner.GlobalContextText <> '', 'PRG_07: Bandeau IHM present');
    ASSERT_FALSE(mainMachine.BusBanner.AlarmBanner.HasAlarm, 'PRG_07: Aucune alarme bloqueuse');
END_TEST

TEST 'MAIN_GLOBAL : Coupure Puissance AU Propagee a tous les Actionneurs'
    // Stimulus : Chute de la boucle AU physique
    mainMachine(
        JoyRawX := 0,
        JoyRawY := 1000,
        JoyDeadmanBtn := TRUE,
        CmdMode := E_Mode.MAINT_N1,
        EmergencyChainClosed := FALSE, // Chaîne AU ouverte
        PowerContactorEngaged := FALSE
    );

    // Vérification : toutes les sorties physiques sont instantanément coupées
    ASSERT_FALSE(mainMachine.BusOutputs.M1RelayFwd, 'Coupure immediate relais M1');
    ASSERT_FALSE(mainMachine.BusOutputs.M1BrakeCmd, 'Frein M1 retombe');
    ASSERT_FALSE(mainMachine.BusOutputs.TranslationBrakeCmd, 'Frein M3 bloque');
END_TEST

TEST 'MAIN_GLOBAL : Relachement homme-mort en contexte cycle -> etape sequencage maintenue (T169-A S3, diag e2e)'
    // ⚠️ Portée honnête : ce test observe la STABILITÉ DU SÉQUENCEUR via l'exposition diag e2e
    // (CycleStep/CycleBusy = sorties réelles de FB_Cycle). Il NE prétend PAS prouver la
    // neutralisation actionneur : dans le mégabloc, le bus vers PRG_04 est alimenté par
    // SeqReq* (entrées externes), pas par les sorties WinchM1Cmd de FB_Cycle. L'invariant
    // « relâchement coupe les demandes actionneur + maintien d'étape » est couvert au niveau
    // unitaire FB_Cycle (TC-P04-020). Ici on vérifie la part réellement tracable e2e.
    // 1. Armement homme-mort + passage Semi-Auto : le séquenceur FB_Cycle quitte X0
    mainMachine(
        JoyRawX := 5000, JoyRawY := 5000, JoyDeadmanBtn := FALSE,
        CmdMode := E_Mode.SEMI_AUTO, CmdWinchSelect := 1,
        EmergencyChainClosed := TRUE, PowerContactorEngaged := TRUE
    );
    mainMachine(
        JoyRawX := 5000, JoyRawY := 5000, JoyDeadmanBtn := TRUE,
        CmdMode := E_Mode.SEMI_AUTO, CmdWinchSelect := 1,
        EmergencyChainClosed := TRUE, PowerContactorEngaged := TRUE
    );
    ADVANCE_TIME(150000000); // > 100 ms DeadmanArmHoldTime
    mainMachine(
        JoyRawX := 5000, JoyRawY := 8000, JoyDeadmanBtn := TRUE,
        CmdMode := E_Mode.SEMI_AUTO, CmdWinchSelect := 1,
        EmergencyChainClosed := TRUE, PowerContactorEngaged := TRUE
    );
    mainMachine(
        JoyRawX := 5000, JoyRawY := 8000, JoyDeadmanBtn := TRUE,
        CmdMode := E_Mode.SEMI_AUTO, CmdWinchSelect := 1,
        EmergencyChainClosed := TRUE, PowerContactorEngaged := TRUE
    );

    // 2. Le séquenceur est observé actif (diag e2e) et le mode arbitre est SEMI_AUTO
    ASSERT_TRUE(mainMachine.CycleStep <> E_AutoCycleStep.AX0_REPOS, 'Sequenceur sorti de X0 en Semi-Auto');
    ASSERT_TRUE(mainMachine.CycleBusy, 'Sequenceur actif (CycleBusy) en Semi-Auto');
    ASSERT_TRUE(mainMachine.BusModes.Mode = E_Mode.SEMI_AUTO, 'Mode SEMI_AUTO arbitre');
    stepBefore := mainMachine.CycleStep;   // mémorise l'étape avant relâchement

    // 3. Relâchement homme-mort / manche au neutre ; X1->X2 avance légitimement (Homed=T par
    //    défaut), donc on n'asserte PAS l'égalité stricte de l'étape. L'invariant e2e réel est
    //    « pas de retour X0 / pas de redémarrage automatique ». Le maintien fin d'étape est
    //    couvert au niveau unitaire FB_Cycle (TC-P04-020).
    mainMachine(
        JoyRawX := 5000, JoyRawY := 5000, JoyDeadmanBtn := FALSE,
        CmdMode := E_Mode.SEMI_AUTO, CmdWinchSelect := 1,
        EmergencyChainClosed := TRUE, PowerContactorEngaged := TRUE
    );
    mainMachine(
        JoyRawX := 5000, JoyRawY := 5000, JoyDeadmanBtn := FALSE,
        CmdMode := E_Mode.SEMI_AUTO, CmdWinchSelect := 1,
        EmergencyChainClosed := TRUE, PowerContactorEngaged := TRUE
    );

    // 4. Pas de retour X0 ni de redémarrage auto au relâchement : l'étape reste « active »
    ASSERT_TRUE(mainMachine.CycleStep <> E_AutoCycleStep.AX0_REPOS, 'Pas de retour X0 au relache (pas de redemarrage auto)');
    ASSERT_TRUE(mainMachine.CycleStep <> E_AutoCycleStep.AX1_INIT OR stepBefore = E_AutoCycleStep.AX0_REPOS,
                'Pas de regression vers le demarrage de cycle');
END_TEST

(* ---- PRG_02_Acquisition_Archi_test.st ---- *)
(* =======================================================================
   🧪 test_prg02_acquisition_archi.st — Architecture PRG_02_Acquisition (TC-P02-001..005)
   ───────────────────────────────────────────────────────────────
   Lot : écriture de tests CI — domaine AF-02 (architecture programme).
   Fiche : DOC/AF/AF_Partie-02_Architecture_Programme_v3.2.md §1 (table des points
           de validation) + AF_Fiche_PRG_02_Acquisition_v1.0.md.
   Conventions : 1 appel harness() = 1 scan ; ADVANCE_TIME(ns) entre les scans pour
   les fronts R_TRIG. Les TC-P02 sont des TC d'architecture : les scénarios valident
   ce qui est testable en boîte noire (population/initialisation/interfaces via
   assertions sur les instances Data/HwIn du harnais) ; les TC de pure architecture
   portent une assertion d'invariant structurel documenté + commentaire
   « (essai d'architecture — validation partielle boîte noire) ».
   ======================================================================= *)

SETUP
VAR
    harness : FB_TestHarness_PRG_02;
END_VAR
END_SETUP

TEST 'TC-P02-001 Un seul producteur par donnee : bus Data qualifie et complet (essai d architecture - validation partielle boite noire)'
    (* Architecture F02.03 : chaque image/bus/commande a un proprietaire unique. En boite
       noire, on verifie que PRG_02 (via le harnais) peuple le bus Data de facon coherente
       et complete : diagnostics DI, qualification codeurs, mesures. *)
    harness(COD1_PosValue := 1008192, COD2_PosValue := 1008192);
    ADVANCE_TIME(10000000);
    harness(COD1_PosValue := 1008192, COD2_PosValue := 1008192);
    ASSERT_TRUE(harness.Data.InputModules.LocalDigitalIoOk, 'Diagnostic module LocalDigitalIoOk publie (producteur unique)');
    ASSERT_TRUE(harness.Data.InputModules.Vh0800EndOk, 'Diagnostic module VH0800 publie');
    ASSERT_TRUE(harness.Data.InputModules.Vh0808EtpOk, 'Diagnostic module VH0808 publie');
    ASSERT_FALSE(harness.Data.InputModules.Fault, 'Pas de defaut module E/S (nominal)');
    ASSERT_TRUE(harness.Data.EncoderM1.Homed, 'Codeur M1 qualifie publie');
    ASSERT_EQ(harness.Data.EncoderM1.Measurement.CablePosM, 2.0, 'Mesure cable M1 publiee (2.0 m)');
END_TEST

TEST 'TC-P02-002 Orchestration ST sans logique cachee : qualification joystick et codeurs (essai d architecture - validation partielle boite noire)'
    (* Architecture F02.02 : les calculs resident dans les FB, le PRG orchestre. En boite
       noire, on verifie que le bus Data porte les resultats qualifies des sous-FB
       (joystick, codeurs) — preuve que l orchestration ST rend les flux lisibles. *)
    harness(JoyRawX := 5000, JoyRawY := 5000, JoyBtnRaw := FALSE);
    ADVANCE_TIME(60000000);
    harness(JoyRawX := 5000, JoyRawY := 5000, JoyBtnRaw := TRUE);
    ADVANCE_TIME(150000000);
    harness(JoyRawX := 5000, JoyRawY := 5000, JoyBtnRaw := TRUE);
    ASSERT_TRUE(harness.Data.Joystick.DeadmanArmed, 'Homme-mort arme (qualification joystick)');
    ASSERT_TRUE((harness.Data.Joystick.AxisX.Direction = 0), 'Axe X au neutre');
    ASSERT_EQ(harness.Data.EncoderM1.Measurement.CablePosM, 2.0, 'Mesure codeur M1 publiee');
END_TEST

TEST 'TC-P02-003 Sorties physiques via PRG_06 : PRG_02 ne produit aucune commande actionneur (essai d architecture - validation partielle boite noire)'
    (* Architecture F02.04 : seul PRG_06_Outputs ecrit les Q/PDO. Le harnais PRG_02 n expose
       que Data (bus) et HwIn (image) — aucune sortie physique. On verifie que l image HwIn
       est bien peuplee (frontiere acquisition) sans commande actionneur. *)
    harness(M1_RelayFwd := TRUE, M1_BrakeCmd := TRUE);
    ADVANCE_TIME(10000000);
    harness(M1_RelayFwd := TRUE, M1_BrakeCmd := TRUE);
    ASSERT_TRUE(harness.HwIn.Winch.M1_ContactorsReleased_DI, 'Image HwIn peuplee (frontiere acquisition)');
    ASSERT_TRUE(harness.HwIn.Machine.PowerContactorEngaged_DI, 'Image machine peuplee');
    (* (essai d architecture - validation partielle boite noire) : le harnais PRG_02 n a aucune
       VAR_OUTPUT de commande actionneur (Q/PDO) — la barriere sortie est PRG_06. *)
END_TEST

TEST 'TC-P02-004 Ordre MainTask conforme : HwIn image arbitree reel/simule (essai d architecture - validation partielle boite noire)'
    (* Architecture F02.01/F02.05 : ordre MainTask + retards N-1. En boite noire, on verifie
       l aiguillage reel/simule : hors simulation, HwIn reflete l image reelle (entrees). *)
    harness(SimulationModeActive := FALSE, M1_ContactorsReleased := FALSE, PowerContactorEngaged := FALSE);
    ADVANCE_TIME(10000000);
    harness(SimulationModeActive := FALSE, M1_ContactorsReleased := FALSE, PowerContactorEngaged := FALSE);
    ASSERT_FALSE(harness.HwIn.Winch.M1_ContactorsReleased_DI, 'Hors simulation -> HwIn reflete le reel (M1 contacteurs relaches)');
    ASSERT_FALSE(harness.HwIn.Machine.PowerContactorEngaged_DI, 'Hors simulation -> HwIn reflete le reel (AU non arme)');
END_TEST

TEST 'TC-P02-005 Troubleshooting lecture seule : PRG_02 produit les diagnostics observes (essai d architecture - validation partielle boite noire)'
    (* Architecture F02.06 : la vue troubleshooting observe seulement. PRG_02 produit les faits
       diagnostiques (InputModuleFault, etats modules) consommes par la vue. En boite noire, on
       verifie que ces diagnostics sont publies sur le bus Data. *)
    harness(COD1_PosValue := 1008192, COD2_PosValue := 1008192);
    ADVANCE_TIME(10000000);
    harness(COD1_PosValue := 1008192, COD2_PosValue := 1008192);
    ASSERT_FALSE(harness.Data.InputModules.Fault, 'Diagnostic InputModuleFault publie (FALSE nominal)');
    ASSERT_TRUE(harness.Data.InputModules.LocalDigitalIoOk, 'Diagnostic module LocalDigitalIoOk publie');
    (* (essai d architecture - validation partielle boite noire) : la lecture seule stricte de la
       vue troubleshooting est couverte en AF-14 (TC-P14-TSV-01..05). *)
END_TEST

(* ---- PRG_02_Acquisition_test.st ---- *)
SETUP
VAR
    harness : FB_TestHarness_PRG_02;
END_VAR
END_SETUP

TEST 'PRG_02_Acquisition : Qualification joystick (neutre -> armement -> consigne X)'
    // 1. Initialisation au neutre
    harness(
        JoyRawX := 5000,
        JoyRawY := 5000,
        JoyBtnRaw := FALSE,
        COD1_PosValue := 1008192, // 2.0 m
        COD2_PosValue := 1008192
    );
    ADVANCE_TIME(60000000);
    harness(JoyRawX := 5000, JoyRawY := 5000, JoyBtnRaw := TRUE); // Appui homme-mort au neutre
    ADVANCE_TIME(150000000); // 150 ms (> 100 ms DeadmanArmHoldTime)
    harness(JoyRawX := 5000, JoyRawY := 5000, JoyBtnRaw := TRUE);

    // Vérification de la structure Data (ST_AcquisitionInterPrg)
    ASSERT_TRUE(harness.Data.Joystick.DeadmanArmed, 'Structure Data: Homme-mort arme avec succes');
    ASSERT_EQ(harness.Data.EncoderM1.Measurement.CablePosM, 2.0, 'Structure Data: Position cable M1 = 2.0m');
    ASSERT_TRUE(harness.Data.EncoderM1.HomedAndReliable, 'Structure Data: Codeur M1 fiabilise');

    // 2. Mouvement manche a droite (RawX = 8000)
    harness(JoyRawX := 8000, JoyRawY := 5000, JoyBtnRaw := TRUE);
    ASSERT_EQ(harness.Data.Joystick.AxisX.Direction, 1, 'Sens X positif detecte (Translation Droite)');
    ASSERT_GT(harness.Data.Joystick.AxisX.SpeedTgt, 0.0, 'Consigne de vitesse non nulle transmise sur le bus Data');

    // Vérification de la structure d'image matérielle HwIn (ST_HardwareImage)
    ASSERT_EQ(harness.HwIn.Operator.JoyXRaw_ANA1, 8000, 'Structure HwIn: JoyXRaw_ANA1 transmis');
    ASSERT_TRUE(harness.HwIn.Operator.JoyBtnRaw, 'Structure HwIn: JoyBtnRaw transmis');
END_TEST

(* ---- PRG_03_Modes_Cycle_test.st ---- *)
SETUP
VAR
    harness : FB_TestHarness_PRG_03;
END_VAR
END_SETUP

TEST 'PRG_03_Modes_Cycle : Mode Manuel MAINT_N1 (arbitrage + autorisations unitaires)'
    harness(
        SelMode := E_Mode.MAINT_N1,
        PowerContactorEngaged := TRUE,
        SelJoystickWinch := 1,        // Selection Joystick M1
        TglMaintenanceZoneAccess := TRUE
    );
    // ---- ST_fbModes_Autorisations : arbitrage mode ----
    ASSERT_EQ(harness.Auth.Mode, E_Mode.MAINT_N1, 'Auth.Mode: MAINT_N1 arbitre');
    // SyncEnable actif par defaut en MAINT_N1 (case IHM cochee par defaut TRUE)
    ASSERT_TRUE(harness.Auth.SyncEnable, 'Auth.SyncEnable vrai en N1 par defaut');
    // Pas d inhibition en MAINT_N1 (N2 only)
    ASSERT_FALSE(harness.Auth.InhibitM1, 'Auth.InhibitM1 faux en N1');
    ASSERT_FALSE(harness.Auth.InhibitM2, 'Auth.InhibitM2 faux en N1');
    // Selection Joystick unitaire autorisee en N1
    ASSERT_EQ(harness.Auth.JoystickWinchSelectArbitrated, 1, 'Auth.JoystickWinchSelectArbitrated = 1 (M1) en N1');
    // HomingApproach : MAINT_N2 only -> faux en N1
    ASSERT_FALSE(harness.Auth.HomingApproachEnable, 'Auth.HomingApproachEnable faux en N1 (N2 only)');
    // Cible Translation Maintenance : N1 OU N2 + bit IHM -> vrai ici
    ASSERT_TRUE(harness.Auth.MaintenanceM3TargetEnable, 'Auth.MaintenanceM3TargetEnable vrai (N1 + bit)');
END_TEST

TEST 'PRG_03_Modes_Cycle : Mode MAINT_N2 (inhibitions exclusives + homing + maintenance)'
    harness(
        SelMode := E_Mode.MAINT_N2,
        PowerContactorEngaged := TRUE,
        SelHomingApproachEnable := TRUE,
        TglMaintenanceZoneAccess := TRUE,
        InhibitM1Request := TRUE,   // front inhibition M1
        SelJoystickWinch := 2        // M2
    );
    // ---- Arbitrage ----
    ASSERT_EQ(harness.Auth.Mode, E_Mode.MAINT_N2, 'Auth.Mode MAINT_N2 arbitre');
    // ---- Inhibitions ----
    ASSERT_TRUE(harness.Auth.InhibitM1, 'Auth.InhibitM1 actif en N2 (demande M1)');
    ASSERT_FALSE(harness.Auth.InhibitM2, 'Auth.InhibitM2 inactif (exclusion mutuelle)');
    // ---- HomingApproach (N2 only) ----
    ASSERT_TRUE(harness.Auth.HomingApproachEnable, 'Auth.HomingApproachEnable vrai en N2');
    // ---- Cible Maintenance ----
    ASSERT_TRUE(harness.Auth.MaintenanceM3TargetEnable, 'Auth.MaintenanceM3TargetEnable vrai en N2 + bit');
    // ---- Selection Joystick unitaire ----
    ASSERT_EQ(harness.Auth.JoystickWinchSelectArbitrated, 2, 'Auth.JoystickWinchSelectArbitrated M2 en N2');
END_TEST

TEST 'PRG_03_Modes_Cycle : Exclusion mutuelle inhibition M1/M2 (jamais les deux actives)'
    harness(
        SelMode := E_Mode.MAINT_N2,
        PowerContactorEngaged := TRUE,
        InhibitM1Request := TRUE,
        InhibitM2Request := TRUE
    );
    // Deux demandes montantes simultanees -> un seul front traite (M1 prioritaire au 1er scan),
    // l autre est rejete. Garantie de securite : JAMAIS les 2 inhibitions actives a la fois.
    ASSERT_TRUE(harness.Auth.InhibitM1 OR harness.Auth.InhibitM2, 'Exactement une inhibition devenue active');
    ASSERT_FALSE(harness.Auth.InhibitM1 AND harness.Auth.InhibitM2, 'Exclusion mutuelle : les 2 inhibitions jamais simultanees');
END_TEST

TEST 'PRG_03_Modes_Cycle : Defaut codeur - SEMI_AUTO selectionne mais cycle non autorise (T207)'
    harness(
        SelMode := E_Mode.SEMI_AUTO,
        PowerContactorEngaged := TRUE,
        EncoderFaultPresent := TRUE,     // defaut codeur agrege
        HomedM1 := TRUE,
        HomedM2 := TRUE
    );
    // T207 : le defaut codeur ne force plus le repli MAINT_N1 ; le mode reste SEMI_AUTO.
    ASSERT_EQ(harness.Auth.Mode, E_Mode.SEMI_AUTO, 'Auth.Mode reste SEMI_AUTO (T207, pas de repli)');
    // Le cycle ne tourne pas : gate codeur FB_Cycle -> sequenceur non Busy.
    ASSERT_FALSE(harness.CycleBusy, 'Cycle non Busy (gate defaut codeur FB_Cycle)');
END_TEST

TEST 'PRG_03_Modes_Cycle : Mode Semi-Auto nominal (sequenceur active, etape initiale)'
    harness(
        SelMode := E_Mode.SEMI_AUTO,
        PowerContactorEngaged := TRUE,
        EncoderFaultPresent := FALSE,
        HomedM1 := TRUE,
        HomedM2 := TRUE,
        DeadmanArmed := TRUE,
        JoystickDeflected := TRUE,
        HeartbeatIhmOk := TRUE
    );
    ASSERT_EQ(harness.Auth.Mode, E_Mode.SEMI_AUTO, 'Auth.Mode SEMI_AUTO arbitre');
    // Sequenceur de cycle prete (etape initiale de preparation)
    ASSERT_EQ(harness.CycleStep, E_AutoCycleStep.AX0_REPOS, 'Sequenceur a l etape X0_PREPARATION');
    ASSERT_FALSE(harness.CycleBusy, 'Sequenceur non Busy initialement');
    ASSERT_FALSE(harness.CycleError, 'Sequenceur sans erreur');
END_TEST

(* ---- PRG_04_Treuils_Benne_test.st ---- *)
SETUP
VAR
    harness : FB_TestHarness_PRG_04;
    acqData : ST_AcquisitionInterPrg;
    modesAuth : ST_Modes_Autorisations;
END_VAR
END_SETUP

TEST 'PRG_04_Treuils_Benne : Commande Montee M1 via Bus AcqData + ModesAuth'
    // 1. Initialisation au repos pour etablir Enable et passer D18
    modesAuth.Mode := E_Mode.MAINT_N1;
    modesAuth.JoystickWinchSelectArbitrated := 1; // M1
    acqData.EncoderM1.Measurement.EncoderAvailable := TRUE;
    acqData.EncoderM1.Measurement.CablePosM := 2.0;

    // Scan 1 au repos (Enable montant)
    harness(
        AcqData := acqData,
        ModesAuth := modesAuth,
        PowerContactorEngaged := TRUE,
        M1_ContactorsReleased := TRUE
    );

    // 2. Application de la commande montee (Scan 2)
    acqData.Joystick.DeadmanArmed := TRUE;
    acqData.Joystick.AtNeutralXY := FALSE;
    acqData.Joystick.AxisY.Direction := 1;

    harness(
        AcqData := acqData,
        ModesAuth := modesAuth,
        BtnWinchM1Up := TRUE,
        PowerContactorEngaged := TRUE,
        M1_ContactorsReleased := TRUE
    );

    // 3. Verification des demandes produites sur le bus sortant ST_WinchInterPrg
    ASSERT_TRUE(harness.Data.WinchM1FinalInterlockRequest.RequestedRelayFwd, 'ST_WinchInterPrg: Ordre RelayFwd genere vers PRG_06');
    ASSERT_FALSE(harness.Data.WinchM1Safety.SafeStop, 'ST_WinchInterPrg: Aucun SafeStop actif');
    ASSERT_GT(harness.Data.M1LogicRequestSpeedCmd_Pct, 0.0, 'ST_WinchInterPrg: consigne vitesse M1 non nulle en montee');
    ASSERT_TRUE(harness.Data.WinchM1State.RelayFwd, 'ST_WinchInterPrg: WinchM1State.RelayFwd reflete la demande');
END_TEST

TEST 'PRG_04_Treuils_Benne : SafeStop Treuil M1 sur Defaut Codeur (Bus AcqData)'
    modesAuth.Mode := E_Mode.MAINT_N1;
    // Stimulus : Defaut codeur remonte par le bus PRG_02
    acqData.EncoderM1.Measurement.EncoderAvailable := FALSE;

    harness(
        AcqData := acqData,
        ModesAuth := modesAuth,
        PowerContactorEngaged := TRUE
    );
    harness(
        AcqData := acqData,
        ModesAuth := modesAuth,
        PowerContactorEngaged := TRUE
    );

    ASSERT_TRUE(harness.Data.WinchM1Safety.SafeStop, 'ST_WinchInterPrg: SafeStop declenche immediatement sur defaut codeur');
    ASSERT_FALSE(harness.Data.WinchM1FinalInterlockRequest.RequestedRelayFwd, 'Mouvement neutralise sur defaut codeur');
END_TEST

(* ---- PRG_05_Translation_test.st ---- *)
SETUP
VAR
    harness   : FB_TestHarness_PRG_05;
    acqData   : ST_AcquisitionInterPrg;
    modesAuth : ST_Modes_Autorisations;
END_VAR
END_SETUP

TEST 'PRG_05_Translation : Commande Translation Fwd (Joystick X + Hauteur Treuils OK)'
    // 1. Contexte : Mode Manuel N1, Câbles treuils hauts (sécurité interlock hauteur validée)
    modesAuth.Mode := E_Mode.MAINT_N1;

    // 2. Stimulus issu du bus PRG_02 : Joystick armé vers la droite (+X)
    acqData.Joystick.DeadmanArmed := TRUE;
    acqData.Joystick.AxisX.Direction := 1;
    acqData.Joystick.AxisX.SpeedTgt := 75.0;

    // 3. Exécution PRG_05 (Position P2/P1/Maintenance = mot valide 00111, ni butée Trémie ni butée Maintenance)
    harness(
        AcqData := acqData,
        ModesAuth := modesAuth,
        WinchM1CablePosM := 5.0,
        WinchM2CablePosM := 5.0,
        M3_PosTremie_DI := FALSE,
        M3_PosPV_DI := FALSE,
        M3_PosPVP2_DI := TRUE,
        M3_PosP1_DI := TRUE,
        M3_PosMaintenance_DI := TRUE,
        PowerContactorEngaged := TRUE,
        DriveOnline := TRUE,
        DriveOperational := TRUE
    );
    ADVANCE_TIME(1000000000);
    harness(
        AcqData := acqData,
        ModesAuth := modesAuth,
        WinchM1CablePosM := 5.0,
        WinchM2CablePosM := 5.0,
        M3_PosTremie_DI := FALSE,
        M3_PosPV_DI := FALSE,
        M3_PosPVP2_DI := TRUE,
        M3_PosP1_DI := TRUE,
        M3_PosMaintenance_DI := TRUE,
        PowerContactorEngaged := TRUE,
        DriveOnline := TRUE,
        DriveOperational := TRUE
    );
    harness(
        AcqData := acqData,
        ModesAuth := modesAuth,
        WinchM1CablePosM := 5.0,
        WinchM2CablePosM := 5.0,
        M3_PosTremie_DI := FALSE,
        M3_PosPV_DI := FALSE,
        M3_PosPVP2_DI := TRUE,
        M3_PosP1_DI := TRUE,
        M3_PosMaintenance_DI := TRUE,
        PowerContactorEngaged := TRUE,
        DriveOnline := TRUE,
        DriveOperational := TRUE
    );

    // 4. Vérification du bus sortant ST_TranslationInterPrg vers PRG_06
    ASSERT_TRUE(harness.Data.TranslationFinalInterlockRequest.BrakeReleaseRequest, 'Demande desserrage frein M3 generee');
    ASSERT_FALSE(harness.Data.TranslationSafety.SafeStop, 'Aucun SafeStop actif sur translation');
    ASSERT_TRUE(harness.Data.TranslationState.ActiveTremie, 'Sens translation avant arbitre');
    ASSERT_GT(harness.Data.TranslationState.SpeedCmd_Pct, 0.0, 'Consigne vitesse M3 arbitree non nulle');
    ASSERT_NEQ(harness.Data.TranslationFinalInterlockRequest.RequestedDriveControlWord, 16#0000, 'ControlWord variateur active pendant la commande');
END_TEST

TEST 'PRG_05_Translation : Commande Translation Rev (Joystick X negatif)'
    modesAuth.Mode := E_Mode.MAINT_N1;
    acqData.Joystick.DeadmanArmed := TRUE;
    acqData.Joystick.AxisX.Direction := -1;
    acqData.Joystick.AxisX.SpeedTgt := 60.0;

    harness(
        AcqData := acqData,
        ModesAuth := modesAuth,
        WinchM1CablePosM := 5.0,
        WinchM2CablePosM := 5.0,
        M3_PosP1_DI := FALSE,
        M3_PosMaintenance_DI := TRUE,
        PowerContactorEngaged := TRUE,
        DriveOnline := TRUE,
        DriveOperational := TRUE
    );
    ADVANCE_TIME(1000000000);
    harness(
        AcqData := acqData,
        ModesAuth := modesAuth,
        WinchM1CablePosM := 5.0,
        WinchM2CablePosM := 5.0,
        M3_PosP1_DI := FALSE,
        M3_PosMaintenance_DI := TRUE,
        PowerContactorEngaged := TRUE,
        DriveOnline := TRUE,
        DriveOperational := TRUE
    );
    harness(
        AcqData := acqData,
        ModesAuth := modesAuth,
        WinchM1CablePosM := 5.0,
        WinchM2CablePosM := 5.0,
        M3_PosP1_DI := FALSE,
        M3_PosMaintenance_DI := TRUE,
        PowerContactorEngaged := TRUE,
        DriveOnline := TRUE,
        DriveOperational := TRUE
    );
    ASSERT_TRUE(harness.Data.TranslationState.ActiveMaintenance, 'Sens translation arriere arbitre');
    ASSERT_TRUE(harness.Data.TranslationFinalInterlockRequest.BrakeReleaseRequest, 'Frein M3 desserre en arriere');
    ASSERT_FALSE(harness.Data.TranslationSafety.SafeStop, 'Aucun SafeStop en commande arriere nominale');
END_TEST

TEST 'PRG_05_Translation : Interdiction Mouvement Translation si Treuils en Bas'
    // Stimulus : Treuil M1 descendu trop bas (< 2m)
    harness(
        AcqData := acqData,
        ModesAuth := modesAuth,
        WinchM1CablePosM := 0.5,
        WinchM2CablePosM := 5.0,
        PowerContactorEngaged := TRUE
    );

    // Vérification : mouvement bloqué par l'interlock de hauteur
    ASSERT_FALSE(harness.Data.TranslationFinalInterlockRequest.BrakeReleaseRequest, 'Frein reste serre');
    ASSERT_FALSE(harness.Data.TranslationState.ActiveTremie, 'Mouvement interdit');
    ASSERT_FALSE(harness.Data.TranslationState.ActiveMaintenance, 'Mouvement interdit');
END_TEST

TEST 'PRG_05_Translation : FdC Tremie LATCHE - un rebond capteur ne libere pas (guard REX MES 2026-09-04)'
    // REGRESSION : un rebond du capteur de butee Tremie (mot 11111 -> 01111 -> 11111)
    // ne doit JAMAIS liberer le bistable M3_LimitSwitchTremieStable ni reautoriser la
    // translation vers la Tremie. On ne perd la butee QU'EN commandant le sens inverse.
    modesAuth.Mode := E_Mode.MAINT_N1;
    acqData.Joystick.DeadmanArmed := TRUE;
    acqData.Joystick.AxisX.Direction := 0;
    acqData.Joystick.AxisX.SpeedTgt := 0.0;

    // 1. Pont sur la butee Tremie : mot 11111 -> bistable latche
    harness(AcqData := acqData, ModesAuth := modesAuth, WinchM1CablePosM := 5.0, WinchM2CablePosM := 5.0,
        M3_PosTremie_DI := TRUE, M3_PosPV_DI := TRUE, M3_PosPVP2_DI := TRUE, M3_PosP1_DI := TRUE, M3_PosMaintenance_DI := TRUE,
        PowerContactorEngaged := TRUE, DriveOnline := TRUE, DriveOperational := TRUE);
    ADVANCE_TIME(500000000);
    harness(AcqData := acqData, ModesAuth := modesAuth, WinchM1CablePosM := 5.0, WinchM2CablePosM := 5.0,
        M3_PosTremie_DI := TRUE, M3_PosPV_DI := TRUE, M3_PosPVP2_DI := TRUE, M3_PosP1_DI := TRUE, M3_PosMaintenance_DI := TRUE,
        PowerContactorEngaged := TRUE, DriveOnline := TRUE, DriveOperational := TRUE);
    ASSERT_TRUE(harness.Data.TranslationState.LimitSwitchTremie, 'Butee Tremie latchee sur mot 11111');

    // 2. REBOND capteur Tremie : DI tombe 2 scans (mot 01111), AUCUNE commande sens inverse
    harness(AcqData := acqData, ModesAuth := modesAuth, WinchM1CablePosM := 5.0, WinchM2CablePosM := 5.0,
        M3_PosTremie_DI := FALSE, M3_PosPV_DI := TRUE, M3_PosPVP2_DI := TRUE, M3_PosP1_DI := TRUE, M3_PosMaintenance_DI := TRUE,
        PowerContactorEngaged := TRUE, DriveOnline := TRUE, DriveOperational := TRUE);
    harness(AcqData := acqData, ModesAuth := modesAuth, WinchM1CablePosM := 5.0, WinchM2CablePosM := 5.0,
        M3_PosTremie_DI := FALSE, M3_PosPV_DI := TRUE, M3_PosPVP2_DI := TRUE, M3_PosP1_DI := TRUE, M3_PosMaintenance_DI := TRUE,
        PowerContactorEngaged := TRUE, DriveOnline := TRUE, DriveOperational := TRUE);
    ASSERT_TRUE(harness.Data.TranslationState.LimitSwitchTremie, 'Rebond capteur -> butee Tremie RESTE latchee (pas de flicker autorisation)');

    // 3. Capteur revient : toujours latche
    harness(AcqData := acqData, ModesAuth := modesAuth, WinchM1CablePosM := 5.0, WinchM2CablePosM := 5.0,
        M3_PosTremie_DI := TRUE, M3_PosPV_DI := TRUE, M3_PosPVP2_DI := TRUE, M3_PosP1_DI := TRUE, M3_PosMaintenance_DI := TRUE,
        PowerContactorEngaged := TRUE, DriveOnline := TRUE, DriveOperational := TRUE);
    ASSERT_TRUE(harness.Data.TranslationState.LimitSwitchTremie, 'Capteur revenu -> toujours latchee');

    // 4. Commande SENS INVERSE (Maintenance, joystick X negatif) -> liberation legitime
    acqData.Joystick.AxisX.Direction := -1;
    acqData.Joystick.AxisX.SpeedTgt := 50.0;
    harness(AcqData := acqData, ModesAuth := modesAuth, WinchM1CablePosM := 5.0, WinchM2CablePosM := 5.0,
        M3_PosTremie_DI := FALSE, M3_PosPV_DI := TRUE, M3_PosPVP2_DI := TRUE, M3_PosP1_DI := TRUE, M3_PosMaintenance_DI := TRUE,
        PowerContactorEngaged := TRUE, DriveOnline := TRUE, DriveOperational := TRUE);
    harness(AcqData := acqData, ModesAuth := modesAuth, WinchM1CablePosM := 5.0, WinchM2CablePosM := 5.0,
        M3_PosTremie_DI := FALSE, M3_PosPV_DI := TRUE, M3_PosPVP2_DI := TRUE, M3_PosP1_DI := TRUE, M3_PosMaintenance_DI := TRUE,
        PowerContactorEngaged := TRUE, DriveOnline := TRUE, DriveOperational := TRUE);
    ASSERT_FALSE(harness.Data.TranslationState.LimitSwitchTremie, 'Commande sens inverse (Maintenance) -> butee Tremie liberee');
END_TEST

(* ═══════════════════════════════════════════════════════════════════════════
   T345 lot L1 — PRG_05 : mémoire de cible et garde de mode des bypass M3.
   ═══════════════════════════════════════════════════════════════════════════ *)

TEST 'TC-P05-T345-01 (T345-L1) La perte de la demande n efface plus la cible deja qualifiee'
    modesAuth.Mode := E_Mode.MAINT_N1;
    acqData.Joystick.DeadmanArmed := TRUE;
    acqData.Joystick.AxisX.Direction := -1;      // demande vers P1/Maintenance
    acqData.Joystick.AxisX.SpeedTgt := 50.0;

    // Scans 1-3 : commande arriere, capteur P1 atteint (mot 00011) -> jeton P1 -> cible qualifiee
    harness(AcqData := acqData, ModesAuth := modesAuth, WinchM1CablePosM := 5.0, WinchM2CablePosM := 5.0,
        M3_PosP1_DI := TRUE, M3_PosMaintenance_DI := TRUE,
        PowerContactorEngaged := TRUE, DriveOnline := TRUE, DriveOperational := TRUE);
    ADVANCE_TIME(1000000000);
    harness(AcqData := acqData, ModesAuth := modesAuth, WinchM1CablePosM := 5.0, WinchM2CablePosM := 5.0,
        M3_PosP1_DI := TRUE, M3_PosMaintenance_DI := TRUE,
        PowerContactorEngaged := TRUE, DriveOnline := TRUE, DriveOperational := TRUE);
    ADVANCE_TIME(1000000000);
    harness(AcqData := acqData, ModesAuth := modesAuth, WinchM1CablePosM := 5.0, WinchM2CablePosM := 5.0,
        M3_PosP1_DI := TRUE, M3_PosMaintenance_DI := TRUE,
        PowerContactorEngaged := TRUE, DriveOnline := TRUE, DriveOperational := TRUE);
    ASSERT_TRUE(harness.Data.TranslationDone, 'cible P1 qualifiee : debounce 100 ms ecoule');

    // Scan 4 : l operateur relache le joystick (perte de la demande) SANS quitter P1.
    // La cible doit rester portee : sans memoire de cible, la detection d arrivee en cours
    // etait effacee et le verrou d arret de l axe ne pouvait plus s armer.
    acqData.Joystick.AxisX.Direction := 0;
    acqData.Joystick.AxisX.SpeedTgt := 0.0;
    harness(AcqData := acqData, ModesAuth := modesAuth, WinchM1CablePosM := 5.0, WinchM2CablePosM := 5.0,
        M3_PosP1_DI := TRUE, M3_PosMaintenance_DI := TRUE,
        PowerContactorEngaged := TRUE, DriveOnline := TRUE, DriveOperational := TRUE);
    ADVANCE_TIME(1000000000);
    harness(AcqData := acqData, ModesAuth := modesAuth, WinchM1CablePosM := 5.0, WinchM2CablePosM := 5.0,
        M3_PosP1_DI := TRUE, M3_PosMaintenance_DI := TRUE,
        PowerContactorEngaged := TRUE, DriveOnline := TRUE, DriveOperational := TRUE);
    ADVANCE_TIME(1000000000);
    harness(AcqData := acqData, ModesAuth := modesAuth, WinchM1CablePosM := 5.0, WinchM2CablePosM := 5.0,
        M3_PosP1_DI := TRUE, M3_PosMaintenance_DI := TRUE,
        PowerContactorEngaged := TRUE, DriveOnline := TRUE, DriveOperational := TRUE);
    ASSERT_TRUE(harness.Data.TranslationDone, 'demande retiree : la cible P1 reste qualifiee');

    // Scans 7-9 : le chariot repart vers la Tremie, le capteur P2 se re-arme (mot 00111) -> un
    // nouveau point est franchi, le jeton P1 retombe et la cible avec lui (elle n est pas collee).
    harness(AcqData := acqData, ModesAuth := modesAuth, WinchM1CablePosM := 5.0, WinchM2CablePosM := 5.0,
        M3_PosPVP2_DI := TRUE, M3_PosP1_DI := TRUE, M3_PosMaintenance_DI := TRUE,
        PowerContactorEngaged := TRUE, DriveOnline := TRUE, DriveOperational := TRUE);
    ADVANCE_TIME(1000000000);
    harness(AcqData := acqData, ModesAuth := modesAuth, WinchM1CablePosM := 5.0, WinchM2CablePosM := 5.0,
        M3_PosPVP2_DI := TRUE, M3_PosP1_DI := TRUE, M3_PosMaintenance_DI := TRUE,
        PowerContactorEngaged := TRUE, DriveOnline := TRUE, DriveOperational := TRUE);
    ADVANCE_TIME(1000000000);
    harness(AcqData := acqData, ModesAuth := modesAuth, WinchM1CablePosM := 5.0, WinchM2CablePosM := 5.0,
        M3_PosPVP2_DI := TRUE, M3_PosP1_DI := TRUE, M3_PosMaintenance_DI := TRUE,
        PowerContactorEngaged := TRUE, DriveOnline := TRUE, DriveOperational := TRUE);
    ASSERT_FALSE(harness.Data.TranslationDone, 'nouveau point franchi : la cible P1 retombe d elle-meme');
END_TEST

TEST 'TC-P05-T345-02 (T345-L1) Bypass de fin de course M3 consomme uniquement en MAINT_N2'
    acqData.Joystick.DeadmanArmed := TRUE;
    acqData.Joystick.AxisX.Direction := 1;       // demande vers la Tremie
    acqData.Joystick.AxisX.SpeedTgt := 50.0;
    modesAuth.Mode := E_Mode.MAINT_N1;           // hors MAINT_N2 : la garde doit s opposer au bypass

    // Scans 1-4 (1 s chacun) : butee Tremie atteinte en demandant (mot 11111), bypass IHM a TRUE et
    // rotation reelle injectee. Hors MAINT_N2 le bypass n est PAS consomme : les deux voies de la
    // cause 6 (axe et safety) doivent s armer, la butee ne peut plus etre neutralisee.
    harness(AcqData := acqData, ModesAuth := modesAuth, WinchM1CablePosM := 5.0, WinchM2CablePosM := 5.0,
        M3_PosTremie_DI := TRUE, M3_PosPV_DI := TRUE, M3_PosPVP2_DI := TRUE, M3_PosP1_DI := TRUE, M3_PosMaintenance_DI := TRUE,
        BypassLimitSwitchIHM := TRUE, DriveActualFreqHzOverride := 5.0,
        PowerContactorEngaged := TRUE, DriveOnline := TRUE, DriveOperational := TRUE);
    ADVANCE_TIME(1000000000);
    harness(AcqData := acqData, ModesAuth := modesAuth, WinchM1CablePosM := 5.0, WinchM2CablePosM := 5.0,
        M3_PosTremie_DI := TRUE, M3_PosPV_DI := TRUE, M3_PosPVP2_DI := TRUE, M3_PosP1_DI := TRUE, M3_PosMaintenance_DI := TRUE,
        BypassLimitSwitchIHM := TRUE, DriveActualFreqHzOverride := 5.0,
        PowerContactorEngaged := TRUE, DriveOnline := TRUE, DriveOperational := TRUE);
    ADVANCE_TIME(1000000000);
    harness(AcqData := acqData, ModesAuth := modesAuth, WinchM1CablePosM := 5.0, WinchM2CablePosM := 5.0,
        M3_PosTremie_DI := TRUE, M3_PosPV_DI := TRUE, M3_PosPVP2_DI := TRUE, M3_PosP1_DI := TRUE, M3_PosMaintenance_DI := TRUE,
        BypassLimitSwitchIHM := TRUE, DriveActualFreqHzOverride := 5.0,
        PowerContactorEngaged := TRUE, DriveOnline := TRUE, DriveOperational := TRUE);
    ADVANCE_TIME(1000000000);
    harness(AcqData := acqData, ModesAuth := modesAuth, WinchM1CablePosM := 5.0, WinchM2CablePosM := 5.0,
        M3_PosTremie_DI := TRUE, M3_PosPV_DI := TRUE, M3_PosPVP2_DI := TRUE, M3_PosP1_DI := TRUE, M3_PosMaintenance_DI := TRUE,
        BypassLimitSwitchIHM := TRUE, DriveActualFreqHzOverride := 5.0,
        PowerContactorEngaged := TRUE, DriveOnline := TRUE, DriveOperational := TRUE);
    ASSERT_TRUE(harness.Data.TranslationState.Error, 'hors MAINT_N2 : cause 6 de l axe NON neutralisee par le bypass');
    ASSERT_TRUE(harness.Data.TranslationSafety.PowerCutOff, 'hors MAINT_N2 : cause 6 safety NON neutralisee -> PowerCutOff');

    // Scans 5-9 : retour en MAINT_N2, meme bypass et memes capteurs -> le bypass est consomme.
    modesAuth.Mode := E_Mode.MAINT_N2;
    harness(AcqData := acqData, ModesAuth := modesAuth, WinchM1CablePosM := 5.0, WinchM2CablePosM := 5.0,
        M3_PosTremie_DI := TRUE, M3_PosPV_DI := TRUE, M3_PosPVP2_DI := TRUE, M3_PosP1_DI := TRUE, M3_PosMaintenance_DI := TRUE,
        BypassLimitSwitchIHM := TRUE, DriveActualFreqHzOverride := 5.0,
        PowerContactorEngaged := TRUE, DriveOnline := TRUE, DriveOperational := TRUE);
    ADVANCE_TIME(1000000000);
    harness(AcqData := acqData, ModesAuth := modesAuth, WinchM1CablePosM := 5.0, WinchM2CablePosM := 5.0,
        M3_PosTremie_DI := TRUE, M3_PosPV_DI := TRUE, M3_PosPVP2_DI := TRUE, M3_PosP1_DI := TRUE, M3_PosMaintenance_DI := TRUE,
        BypassLimitSwitchIHM := TRUE, DriveActualFreqHzOverride := 5.0,
        PowerContactorEngaged := TRUE, DriveOnline := TRUE, DriveOperational := TRUE);
    ADVANCE_TIME(1000000000);
    harness(AcqData := acqData, ModesAuth := modesAuth, WinchM1CablePosM := 5.0, WinchM2CablePosM := 5.0,
        M3_PosTremie_DI := TRUE, M3_PosPV_DI := TRUE, M3_PosPVP2_DI := TRUE, M3_PosP1_DI := TRUE, M3_PosMaintenance_DI := TRUE,
        BypassLimitSwitchIHM := TRUE, DriveActualFreqHzOverride := 5.0,
        PowerContactorEngaged := TRUE, DriveOnline := TRUE, DriveOperational := TRUE);
    ADVANCE_TIME(1000000000);
    harness(AcqData := acqData, ModesAuth := modesAuth, WinchM1CablePosM := 5.0, WinchM2CablePosM := 5.0,
        M3_PosTremie_DI := TRUE, M3_PosPV_DI := TRUE, M3_PosPVP2_DI := TRUE, M3_PosP1_DI := TRUE, M3_PosMaintenance_DI := TRUE,
        BypassLimitSwitchIHM := TRUE, DriveActualFreqHzOverride := 5.0,
        PowerContactorEngaged := TRUE, DriveOnline := TRUE, DriveOperational := TRUE);
    ADVANCE_TIME(1000000000);
    harness(AcqData := acqData, ModesAuth := modesAuth, WinchM1CablePosM := 5.0, WinchM2CablePosM := 5.0,
        M3_PosTremie_DI := TRUE, M3_PosPV_DI := TRUE, M3_PosPVP2_DI := TRUE, M3_PosP1_DI := TRUE, M3_PosMaintenance_DI := TRUE,
        BypassLimitSwitchIHM := TRUE, DriveActualFreqHzOverride := 5.0,
        PowerContactorEngaged := TRUE, DriveOnline := TRUE, DriveOperational := TRUE);
    ASSERT_FALSE(harness.Data.TranslationState.Error, 'en MAINT_N2 : bypass consomme -> cause 6 de l axe neutralisee');
    ASSERT_FALSE(harness.Data.TranslationSafety.PowerCutOff, 'en MAINT_N2 : bypass consomme -> pas de PowerCutOff');
END_TEST

(* ---- PRG_06_Outputs_test.st ---- *)
SETUP
VAR
    harness         : FB_TestHarness_PRG_06;
    winchData       : ST_WinchInterPrg;
    translationData : ST_TranslationInterPrg;
END_VAR
END_SETUP

TEST 'PRG_06_Outputs : Transmission Ordres M1 et M3 en Marche Normale'
    // 1. Contexte M1 : Demande de montee active palier 1
    winchData.WinchM1FinalInterlockRequest.Enable := TRUE;
    winchData.WinchM1FinalInterlockRequest.PowerContactorEngaged := TRUE;
    winchData.WinchM1FinalInterlockRequest.SafeStop := FALSE;
    winchData.WinchM1FinalInterlockRequest.PowerCutOff := FALSE;
    winchData.WinchM1FinalInterlockRequest.AscentPermit := TRUE;
    winchData.WinchM1FinalInterlockRequest.DescendPermit := TRUE;
    winchData.WinchM1FinalInterlockRequest.BrakeFeedback := TRUE;
    winchData.WinchM1FinalInterlockRequest.FwdRevSpeedFeedbackOff := TRUE;
    winchData.WinchM1FinalInterlockRequest.RequestedRelayFwd := TRUE;
    winchData.WinchM1FinalInterlockRequest.RequestedRelayRev := FALSE;
    winchData.WinchM1FinalInterlockRequest.RequestedContactor1 := FALSE;
    winchData.WinchM1FinalInterlockRequest.RequestedStep := 1;

    // 2. Contexte M3 : Demande de frein relache
    translationData.TranslationFinalInterlockRequest.Enable := TRUE;
    translationData.TranslationFinalInterlockRequest.PowerContactorEngaged := TRUE;
    translationData.TranslationFinalInterlockRequest.SafeStop := FALSE;
    translationData.TranslationFinalInterlockRequest.PowerCutOff := FALSE;
    translationData.TranslationFinalInterlockRequest.BrakeReleaseRequest := TRUE;

    harness(WinchData := winchData, TranslationData := translationData);

    // 3. Verification des sorties reelles sur le bus ST_OutputsInterPrg
    ASSERT_TRUE(harness.Data.M1RelayFwd, 'Contacteur montee M1 active');
    ASSERT_TRUE(harness.Data.M1BrakeCmd, 'Commande desserrage frein M1 active');
    ASSERT_TRUE(harness.Data.TranslationBrakeCmd, 'Commande desserrage frein M3 active');
END_TEST

TEST 'PRG_06_Outputs : Transmission Ordre M2 en Marche Normale'
    // Contexte M2 : Demande de montee (fermeture) active palier 1
    winchData.WinchM2FinalInterlockRequest.Enable := TRUE;
    winchData.WinchM2FinalInterlockRequest.PowerContactorEngaged := TRUE;
    winchData.WinchM2FinalInterlockRequest.SafeStop := FALSE;
    winchData.WinchM2FinalInterlockRequest.PowerCutOff := FALSE;
    winchData.WinchM2FinalInterlockRequest.AscentPermit := TRUE;
    winchData.WinchM2FinalInterlockRequest.DescendPermit := TRUE;
    winchData.WinchM2FinalInterlockRequest.BrakeFeedback := TRUE;
    winchData.WinchM2FinalInterlockRequest.FwdRevSpeedFeedbackOff := TRUE;
    winchData.WinchM2FinalInterlockRequest.RequestedRelayFwd := TRUE;
    winchData.WinchM2FinalInterlockRequest.RequestedRelayRev := FALSE;
    winchData.WinchM2FinalInterlockRequest.RequestedContactor1 := FALSE;
    winchData.WinchM2FinalInterlockRequest.RequestedStep := 1;

    harness(WinchData := winchData, TranslationData := translationData);

    // Verification sorties M2
    ASSERT_TRUE(harness.Data.M2RelayFwd, 'Contacteur montee (fermeture) M2 active');
    ASSERT_TRUE(harness.Data.M2BrakeCmd, 'Commande desserrage frein M2 active');
END_TEST

TEST 'PRG_06_Outputs : Barriere de Securite Coupure Brutale PowerCutOff sur M1'
    // Stimulus : Commande active MAIS PowerCutOff = TRUE (Arret d'urgence ou defaut critique)
    winchData.WinchM1FinalInterlockRequest.Enable := TRUE;
    winchData.WinchM1FinalInterlockRequest.PowerContactorEngaged := TRUE;
    winchData.WinchM1FinalInterlockRequest.PowerCutOff := TRUE;
    winchData.WinchM1FinalInterlockRequest.RequestedRelayFwd := TRUE;
    winchData.WinchM1FinalInterlockRequest.RequestedContactor1 := TRUE;
    winchData.WinchM1FinalInterlockRequest.RequestedStep := 1;

    harness(
        WinchData := winchData,
        TranslationData := translationData
    );

    // Verification : barriere infranchissable, toutes sorties a zero
    ASSERT_FALSE(harness.Data.M1RelayFwd, 'Relais montee coupe');
    ASSERT_FALSE(harness.Data.M1SpeedContactor1, 'Contacteur de vitesse coupe');
    ASSERT_FALSE(harness.Data.M1BrakeCmd, 'Frein M1 force a l arret (non desserre)');
END_TEST
